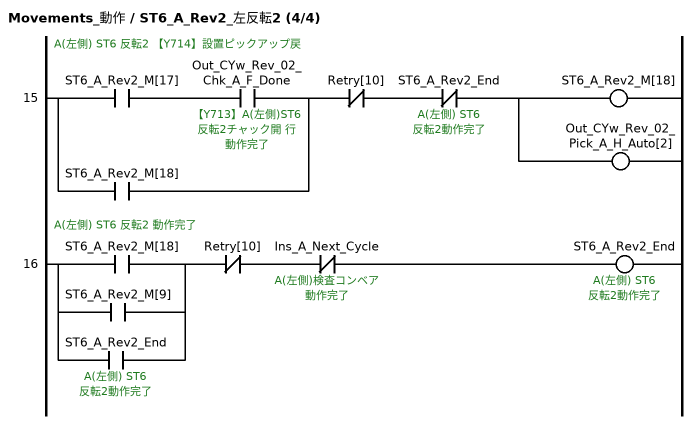
(* [picture p48: Movements_動作 / ST6_A_Rev2_左反転2, rungs 15-16] *)
(* Rung 15: A(左側) ST6 反転2 【Y714】設置ピックアップ戻 *)
_p89 := ((ST6_A_Rev2_M[17] AND Out_CYw_Rev_02_Chk_A_F_Done) OR ST6_A_Rev2_M[18]) AND NOT Retry[10] AND NOT ST6_A_Rev2_End;
ST6_A_Rev2_M[18] := _p89;
Out_CYw_Rev_02_Pick_A_H_Auto[2] := _p89;
(* Rung 16: A(左側) ST6 反転2 動作完了 *)
ST6_A_Rev2_End := (ST6_A_Rev2_M[18] OR ST6_A_Rev2_M[9] OR ST6_A_Rev2_End) AND NOT Retry[10] AND NOT Ins_A_Next_Cycle;

(* Section ST7_A_Dis2_左SF排出: ladder, written here as Structured Text *)

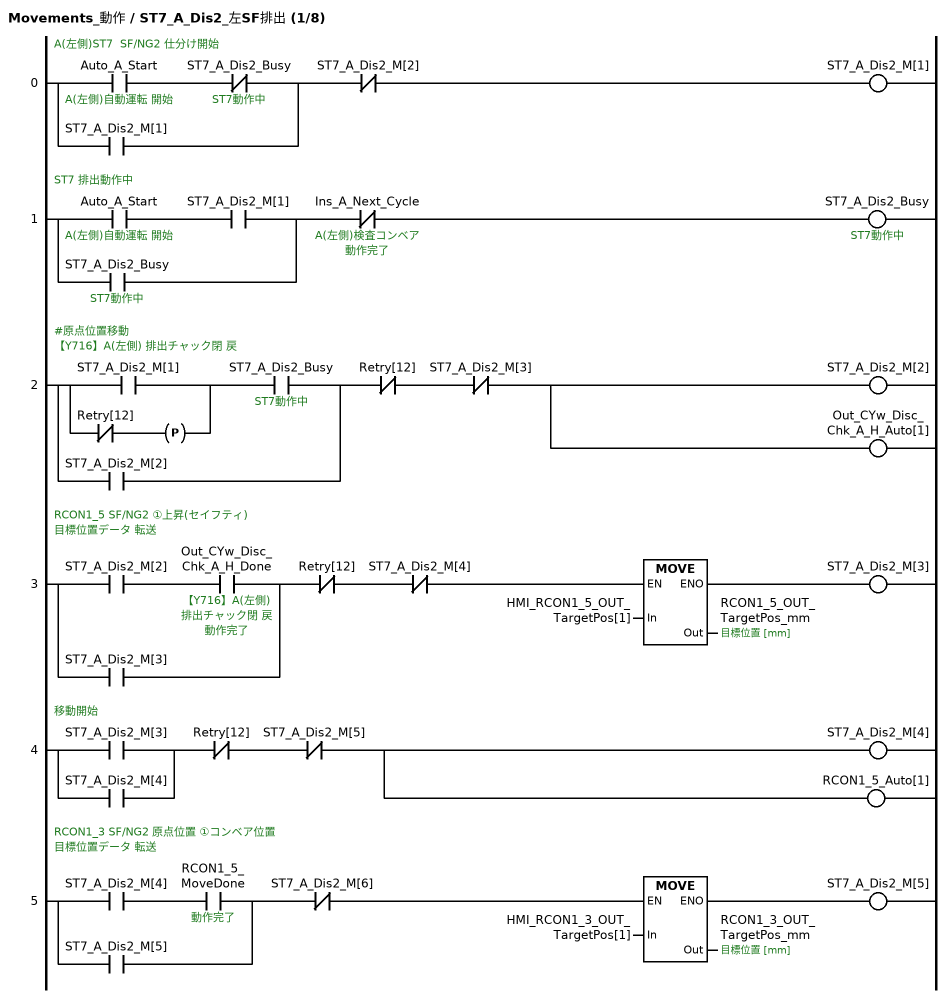
(* Rung 0: A(左側)ST7  SF/NG2 仕分け開始 *)
ST7_A_Dis2_M[1] := ((Auto_A_Start AND NOT ST7_A_Dis2_Busy) OR ST7_A_Dis2_M[1]) AND NOT ST7_A_Dis2_M[2];
(* Rung 1: ST7 排出動作中 *)
ST7_A_Dis2_Busy := ((Auto_A_Start AND ST7_A_Dis2_M[1]) OR ST7_A_Dis2_Busy) AND NOT Ins_A_Next_Cycle;
(* Rung 2: #原点位置移動 / 【Y716】A(左側) 排出チャック閉 戻 *)
_e90(CLK := NOT Retry[12]);
_p91 := (((ST7_A_Dis2_M[1] OR _e90.Q) AND ST7_A_Dis2_Busy) OR ST7_A_Dis2_M[2]) AND NOT Retry[12] AND NOT ST7_A_Dis2_M[3];
ST7_A_Dis2_M[2] := _p91;
Out_CYw_Disc_Chk_A_H_Auto[1] := _p91;
(* Rung 3: RCON1_5 SF/NG2 ①上昇(セイフティ) / 目標位置データ 転送 *)
IF ((ST7_A_Dis2_M[2] AND Out_CYw_Disc_Chk_A_H_Done) OR ST7_A_Dis2_M[3]) AND NOT Retry[12] AND NOT ST7_A_Dis2_M[4] THEN
    RCON1_5_OUT_TargetPos_mm := HMI_RCON1_5_OUT_TargetPos[1];
END_IF;
ST7_A_Dis2_M[3] := ((ST7_A_Dis2_M[2] AND Out_CYw_Disc_Chk_A_H_Done) OR ST7_A_Dis2_M[3]) AND NOT Retry[12] AND NOT ST7_A_Dis2_M[4];
(* Rung 4: 移動開始 *)
_p92 := (ST7_A_Dis2_M[3] OR ST7_A_Dis2_M[4]) AND NOT Retry[12] AND NOT ST7_A_Dis2_M[5];
ST7_A_Dis2_M[4] := _p92;
RCON1_5_Auto[1] := _p92;
(* Rung 5: RCON1_3 SF/NG2 原点位置 ①コンベア位置 / 目標位置データ 転送 *)
IF ((ST7_A_Dis2_M[4] AND RCON1_5_MoveDone) OR ST7_A_Dis2_M[5]) AND NOT ST7_A_Dis2_M[6] THEN
    RCON1_3_OUT_TargetPos_mm := HMI_RCON1_3_OUT_TargetPos[1];
END_IF;
ST7_A_Dis2_M[5] := ((ST7_A_Dis2_M[4] AND RCON1_5_MoveDone) OR ST7_A_Dis2_M[5]) AND NOT ST7_A_Dis2_M[6];

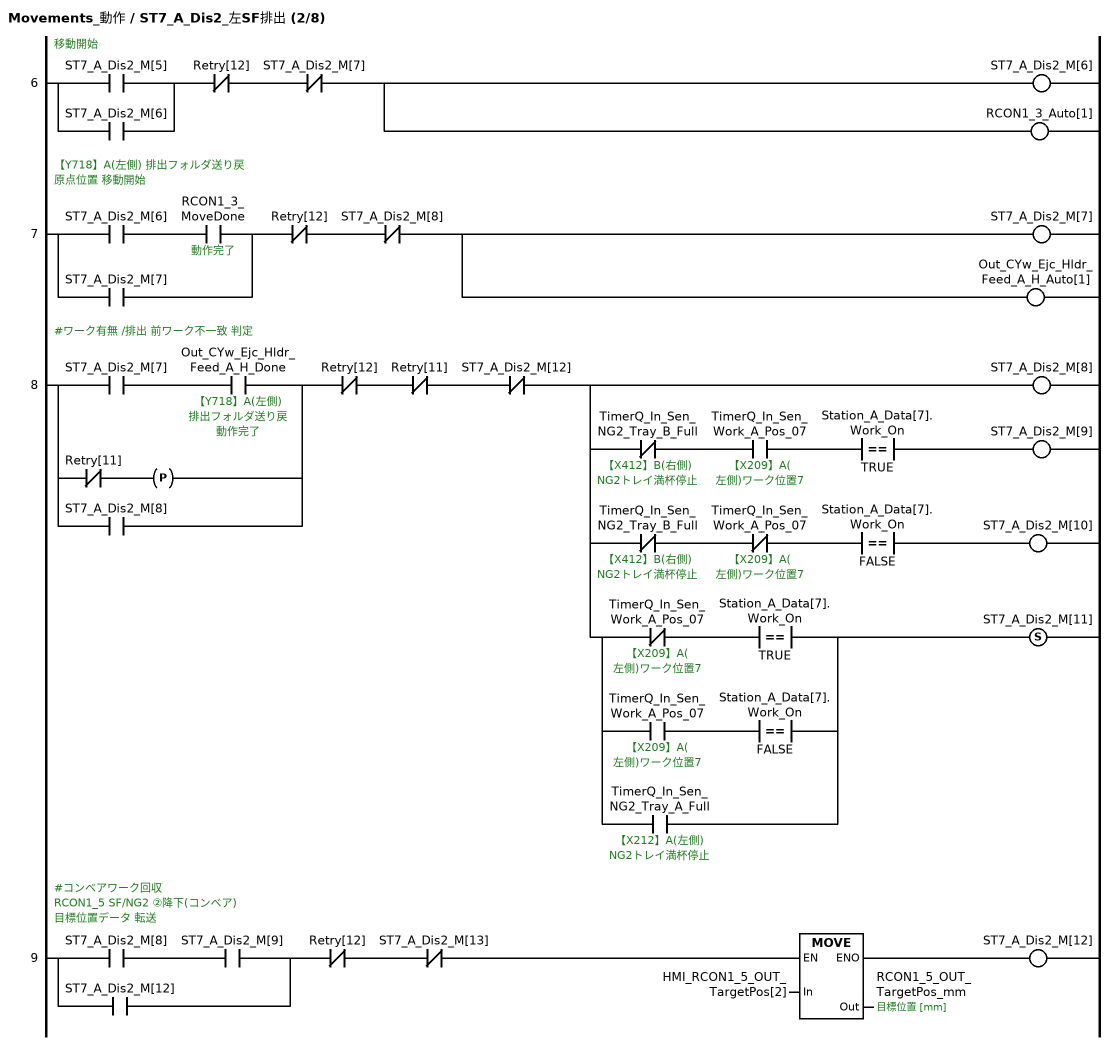
(* Rung 6: 移動開始 *)
_p93 := (ST7_A_Dis2_M[5] OR ST7_A_Dis2_M[6]) AND NOT Retry[12] AND NOT ST7_A_Dis2_M[7];
ST7_A_Dis2_M[6] := _p93;
RCON1_3_Auto[1] := _p93;
(* Rung 7: 【Y718】A(左側) 排出フォルダ送り戻 / 原点位置 移動開始 *)
_p94 := ((ST7_A_Dis2_M[6] AND RCON1_3_MoveDone) OR ST7_A_Dis2_M[7]) AND NOT Retry[12] AND NOT ST7_A_Dis2_M[8];
ST7_A_Dis2_M[7] := _p94;
Out_CYw_Ejc_Hldr_Feed_A_H_Auto[1] := _p94;
(* Rung 8: #ワーク有無 /排出 前ワーク不一致 判定 *)
_e95(CLK := NOT Retry[11]);
_p96 := ((ST7_A_Dis2_M[7] AND Out_CYw_Ejc_Hldr_Feed_A_H_Done) OR _e95.Q OR ST7_A_Dis2_M[8]) AND NOT Retry[12] AND NOT Retry[11] AND NOT ST7_A_Dis2_M[12];
ST7_A_Dis2_M[8] := _p96;
ST7_A_Dis2_M[9] := _p96 AND NOT TimerQ_In_Sen_NG2_Tray_B_Full AND TimerQ_In_Sen_Work_A_Pos_07 AND (Station_A_Data[7].Work_On = TRUE);
ST7_A_Dis2_M[10] := _p96 AND NOT TimerQ_In_Sen_NG2_Tray_B_Full AND NOT TimerQ_In_Sen_Work_A_Pos_07 AND (Station_A_Data[7].Work_On = FALSE);
IF _p96 AND ((NOT TimerQ_In_Sen_Work_A_Pos_07 AND (Station_A_Data[7].Work_On = TRUE)) OR (TimerQ_In_Sen_Work_A_Pos_07 AND (Station_A_Data[7].Work_On = FALSE)) OR TimerQ_In_Sen_NG2_Tray_A_Full) THEN
    ST7_A_Dis2_M[11] := TRUE;
END_IF;
(* Rung 9: #コンベアワーク回収 / RCON1_5 SF/NG2 ②降下(コンベア) / 目標位置データ 転送 *)
IF ((ST7_A_Dis2_M[8] AND ST7_A_Dis2_M[9]) OR ST7_A_Dis2_M[12]) AND NOT Retry[12] AND NOT ST7_A_Dis2_M[13] THEN
    RCON1_5_OUT_TargetPos_mm := HMI_RCON1_5_OUT_TargetPos[2];
END_IF;
ST7_A_Dis2_M[12] := ((ST7_A_Dis2_M[8] AND ST7_A_Dis2_M[9]) OR ST7_A_Dis2_M[12]) AND NOT Retry[12] AND NOT ST7_A_Dis2_M[13];

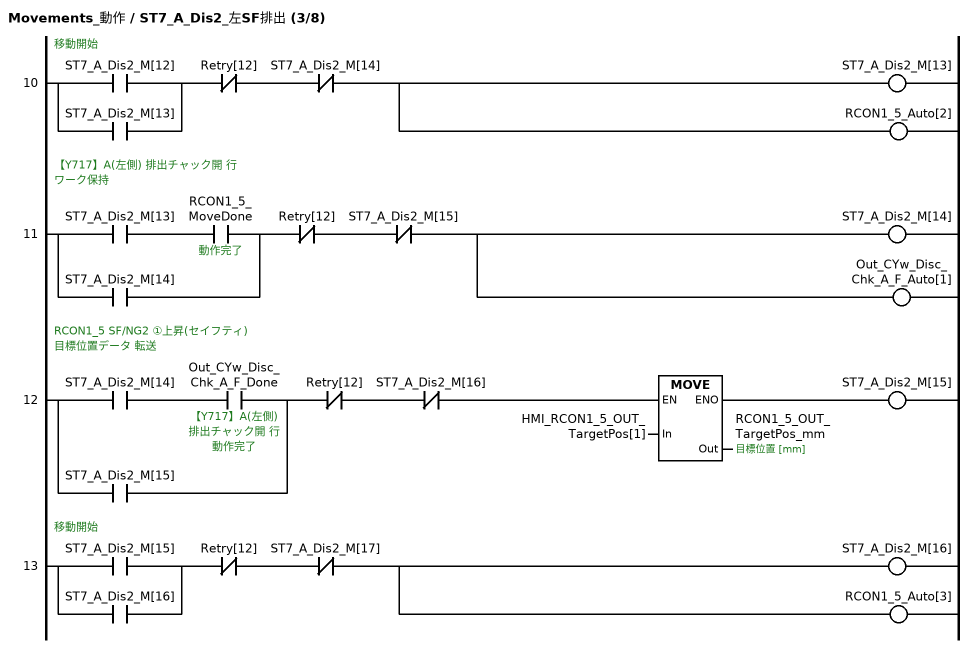
(* Rung 10: 移動開始 *)
_p97 := (ST7_A_Dis2_M[12] OR ST7_A_Dis2_M[13]) AND NOT Retry[12] AND NOT ST7_A_Dis2_M[14];
ST7_A_Dis2_M[13] := _p97;
RCON1_5_Auto[2] := _p97;
(* Rung 11: 【Y717】A(左側) 排出チャック開 行 / ワーク保持 *)
_p98 := ((ST7_A_Dis2_M[13] AND RCON1_5_MoveDone) OR ST7_A_Dis2_M[14]) AND NOT Retry[12] AND NOT ST7_A_Dis2_M[15];
ST7_A_Dis2_M[14] := _p98;
Out_CYw_Disc_Chk_A_F_Auto[1] := _p98;
(* Rung 12: RCON1_5 SF/NG2 ①上昇(セイフティ) / 目標位置データ 転送 *)
IF ((ST7_A_Dis2_M[14] AND Out_CYw_Disc_Chk_A_F_Done) OR ST7_A_Dis2_M[15]) AND NOT Retry[12] AND NOT ST7_A_Dis2_M[16] THEN
    RCON1_5_OUT_TargetPos_mm := HMI_RCON1_5_OUT_TargetPos[1];
END_IF;
ST7_A_Dis2_M[15] := ((ST7_A_Dis2_M[14] AND Out_CYw_Disc_Chk_A_F_Done) OR ST7_A_Dis2_M[15]) AND NOT Retry[12] AND NOT ST7_A_Dis2_M[16];
(* Rung 13: 移動開始 *)
_p99 := (ST7_A_Dis2_M[15] OR ST7_A_Dis2_M[16]) AND NOT Retry[12] AND NOT ST7_A_Dis2_M[17];
ST7_A_Dis2_M[16] := _p99;
RCON1_5_Auto[3] := _p99;

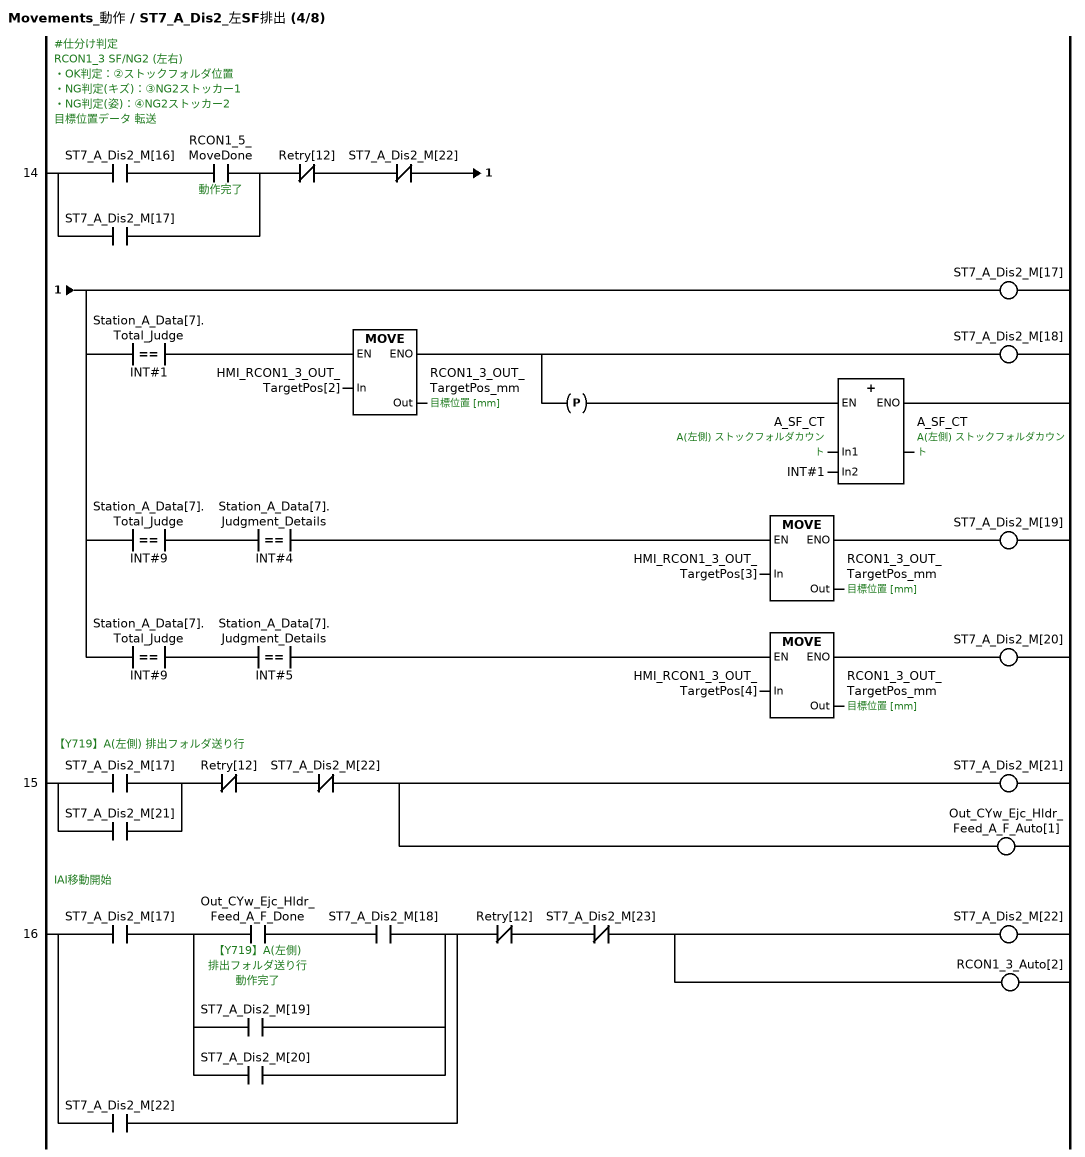
(* Rung 14: #仕分け判定 / RCON1_3 SF/NG2 (左右) / ・OK判定：②ストックフォルダ位置 / ・NG判定(キズ)：③NG2ストッカー1 / ・NG判定(姿)：④NG2ストッカー2 / 目標位置データ 転送 *)
_p100 := ((ST7_A_Dis2_M[16] AND RCON1_5_MoveDone) OR ST7_A_Dis2_M[17]) AND NOT Retry[12] AND NOT ST7_A_Dis2_M[22];
ST7_A_Dis2_M[17] := _p100;
IF _p100 AND (Station_A_Data[7].Total_Judge = INT#1) THEN
    RCON1_3_OUT_TargetPos_mm := HMI_RCON1_3_OUT_TargetPos[2];
END_IF;
_p101 := _p100 AND (Station_A_Data[7].Total_Judge = INT#1);
ST7_A_Dis2_M[18] := _p101;
_e102(CLK := _p101);
IF _e102.Q THEN A_SF_CT := A_SF_CT + INT#1; END_IF;
IF _p100 AND (Station_A_Data[7].Total_Judge = INT#9) AND (Station_A_Data[7].Judgment_Details = INT#4) THEN
    RCON1_3_OUT_TargetPos_mm := HMI_RCON1_3_OUT_TargetPos[3];
END_IF;
ST7_A_Dis2_M[19] := _p100 AND (Station_A_Data[7].Total_Judge = INT#9) AND (Station_A_Data[7].Judgment_Details = INT#4);
IF _p100 AND (Station_A_Data[7].Total_Judge = INT#9) AND (Station_A_Data[7].Judgment_Details = INT#5) THEN
    RCON1_3_OUT_TargetPos_mm := HMI_RCON1_3_OUT_TargetPos[4];
END_IF;
ST7_A_Dis2_M[20] := _p100 AND (Station_A_Data[7].Total_Judge = INT#9) AND (Station_A_Data[7].Judgment_Details = INT#5);
(* Rung 15: 【Y719】A(左側) 排出フォルダ送り行 *)
_p103 := (ST7_A_Dis2_M[17] OR ST7_A_Dis2_M[21]) AND NOT Retry[12] AND NOT ST7_A_Dis2_M[22];
ST7_A_Dis2_M[21] := _p103;
Out_CYw_Ejc_Hldr_Feed_A_F_Auto[1] := _p103;
(* Rung 16: IAI移動開始 *)
_p104 := ((ST7_A_Dis2_M[17] AND ((Out_CYw_Ejc_Hldr_Feed_A_F_Done AND ST7_A_Dis2_M[18]) OR ST7_A_Dis2_M[19] OR ST7_A_Dis2_M[20])) OR ST7_A_Dis2_M[22]) AND NOT Retry[12] AND NOT ST7_A_Dis2_M[23];
ST7_A_Dis2_M[22] := _p104;
RCON1_3_Auto[2] := _p104;

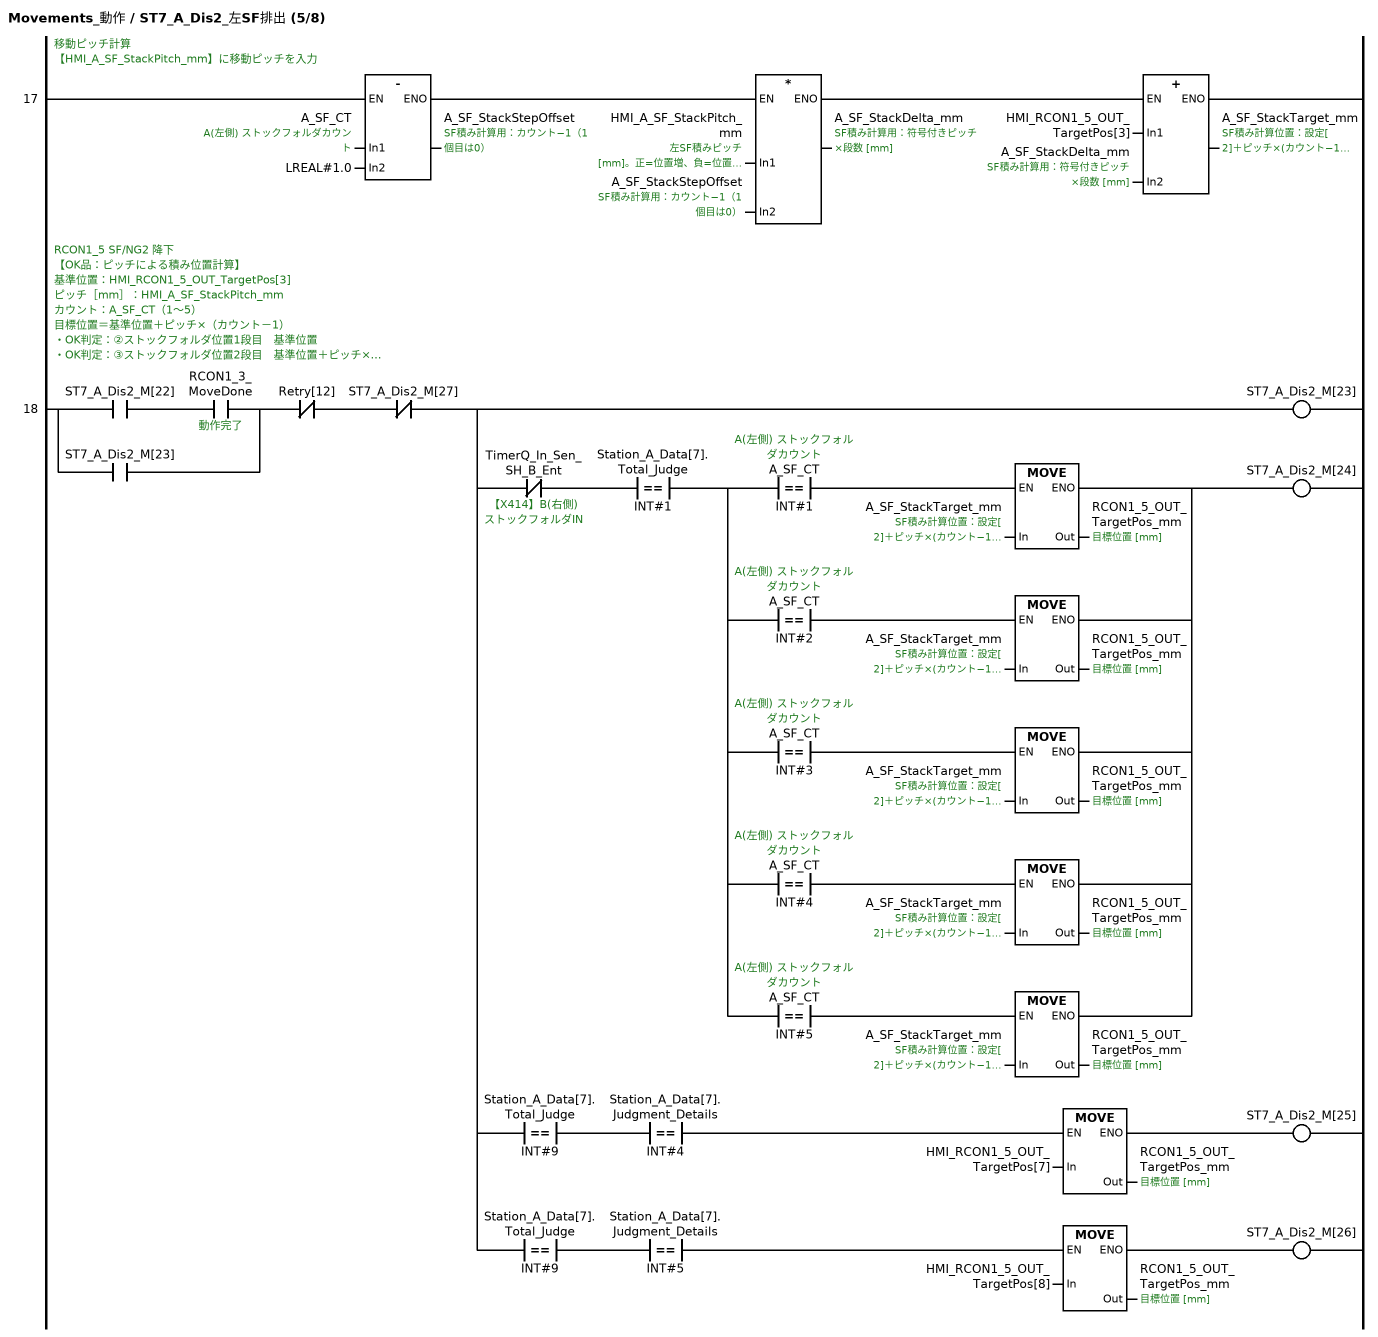
(* Rung 17: 移動ピッチ計算 / 【HMI_A_SF_StackPitch_mm】に移動ピッチを入力 *)
A_SF_StackStepOffset := A_SF_CT - LREAL#1.0;
A_SF_StackDelta_mm := HMI_A_SF_StackPitch_mm * A_SF_StackStepOffset;
A_SF_StackTarget_mm := HMI_RCON1_5_OUT_TargetPos[3] + A_SF_StackDelta_mm;
(* Rung 18: RCON1_5 SF/NG2 降下 / 【OK品：ピッチによる積み位置計算】 / 基準位置：HMI_RCON1_5_OUT_TargetPos[3] / ピッチ［mm］：HMI_A_SF_StackPitch_mm / カウント：A_SF_CT（1～5） / 目標位置＝基準位置＋ピッチ×（カウント－1） / ・OK判定：②ストックフォルダ位置1段目　基準位置 / ・OK判定：③ストックフォルダ位置2段目　基準位置＋ピッチ×1 / ・OK判定：④ストックフォルダ位置3段目　基準位置＋ピッチ×2 / ・OK判定：⑤ストックフォルダ位置4段目　基準位置＋ピッチ×3 / ・OK判定：⑥ストックフォルダ位置5段目　基準位置＋ピッチ×4 / 【NG品：従来の固定位置を使用】 / ・NG判定(キズ)：⑦NG2ストッカー1 / ・NG判定(姿)：⑧NG2ストッカー2 / 目標位置データ 転送 *)
_p105 := ((ST7_A_Dis2_M[22] AND RCON1_3_MoveDone) OR ST7_A_Dis2_M[23]) AND NOT Retry[12] AND NOT ST7_A_Dis2_M[27];
ST7_A_Dis2_M[23] := _p105;
_p106 := _p105 AND NOT TimerQ_In_Sen_SH_B_Ent AND (Station_A_Data[7].Total_Judge = INT#1);
IF _p106 AND (A_SF_CT = INT#1) THEN RCON1_5_OUT_TargetPos_mm := A_SF_StackTarget_mm; END_IF;
IF _p106 AND (A_SF_CT = INT#2) THEN RCON1_5_OUT_TargetPos_mm := A_SF_StackTarget_mm; END_IF;
IF _p106 AND (A_SF_CT = INT#3) THEN RCON1_5_OUT_TargetPos_mm := A_SF_StackTarget_mm; END_IF;
IF _p106 AND (A_SF_CT = INT#4) THEN RCON1_5_OUT_TargetPos_mm := A_SF_StackTarget_mm; END_IF;
IF _p106 AND (A_SF_CT = INT#5) THEN RCON1_5_OUT_TargetPos_mm := A_SF_StackTarget_mm; END_IF;
ST7_A_Dis2_M[24] := _p106 AND ((A_SF_CT = INT#1) OR (A_SF_CT = INT#2) OR (A_SF_CT = INT#3) OR (A_SF_CT = INT#4) OR (A_SF_CT = INT#5));
IF _p105 AND (Station_A_Data[7].Total_Judge = INT#9) AND (Station_A_Data[7].Judgment_Details = INT#4) THEN
    RCON1_5_OUT_TargetPos_mm := HMI_RCON1_5_OUT_TargetPos[7];
END_IF;
ST7_A_Dis2_M[25] := _p105 AND (Station_A_Data[7].Total_Judge = INT#9) AND (Station_A_Data[7].Judgment_Details = INT#4);
IF _p105 AND (Station_A_Data[7].Total_Judge = INT#9) AND (Station_A_Data[7].Judgment_Details = INT#5) THEN
    RCON1_5_OUT_TargetPos_mm := HMI_RCON1_5_OUT_TargetPos[8];
END_IF;
ST7_A_Dis2_M[26] := _p105 AND (Station_A_Data[7].Total_Judge = INT#9) AND (Station_A_Data[7].Judgment_Details = INT#5);

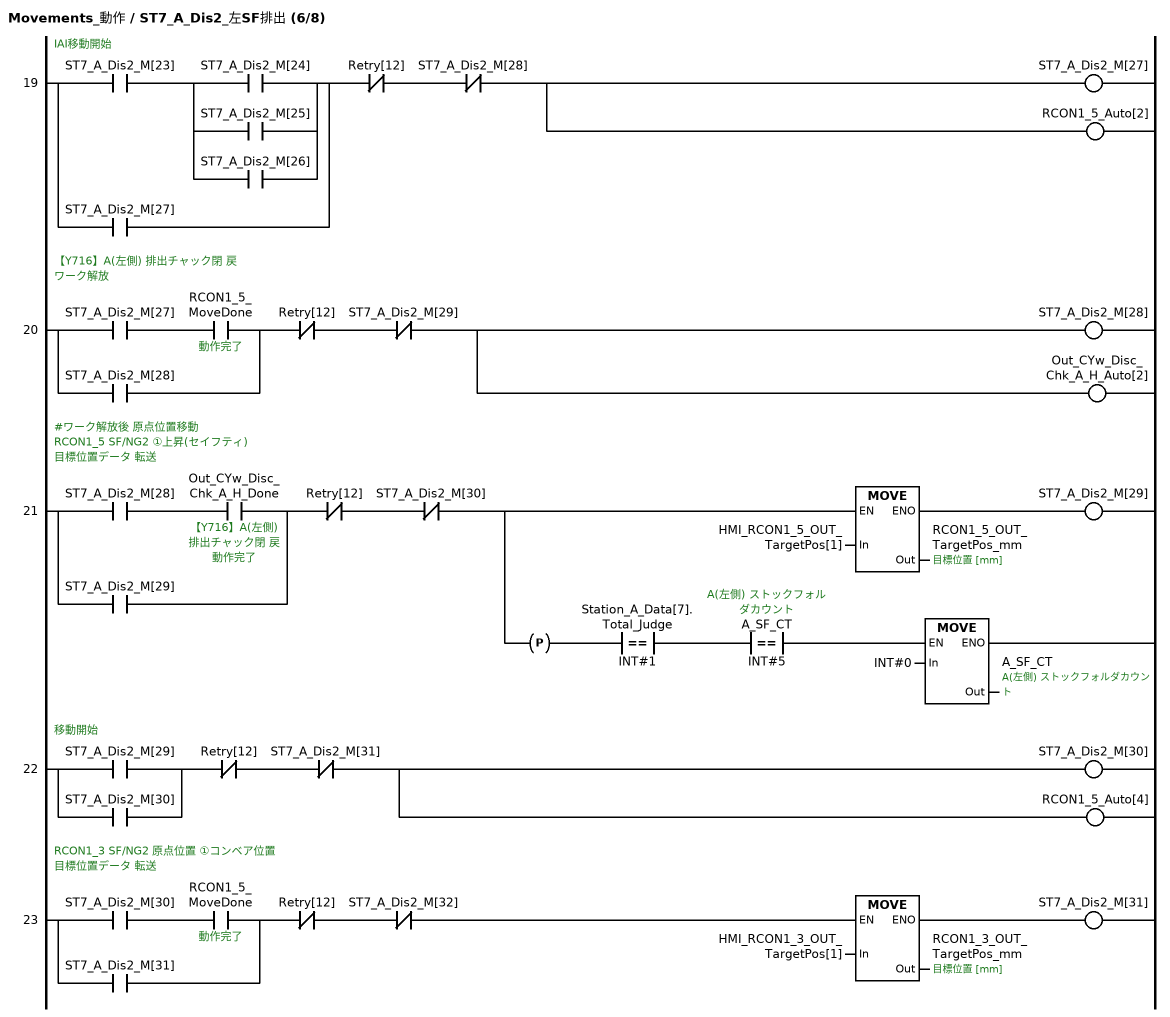
(* Rung 19: IAI移動開始 *)
_p107 := ((ST7_A_Dis2_M[23] AND (ST7_A_Dis2_M[24] OR ST7_A_Dis2_M[25] OR ST7_A_Dis2_M[26])) OR ST7_A_Dis2_M[27]) AND NOT Retry[12] AND NOT ST7_A_Dis2_M[28];
ST7_A_Dis2_M[27] := _p107;
RCON1_5_Auto[2] := _p107;
(* Rung 20: 【Y716】A(左側) 排出チャック閉 戻 / ワーク解放 *)
_p108 := ((ST7_A_Dis2_M[27] AND RCON1_5_MoveDone) OR ST7_A_Dis2_M[28]) AND NOT Retry[12] AND NOT ST7_A_Dis2_M[29];
ST7_A_Dis2_M[28] := _p108;
Out_CYw_Disc_Chk_A_H_Auto[2] := _p108;
(* Rung 21: #ワーク解放後 原点位置移動 / RCON1_5 SF/NG2 ①上昇(セイフティ) / 目標位置データ 転送 *)
_p109 := ((ST7_A_Dis2_M[28] AND Out_CYw_Disc_Chk_A_H_Done) OR ST7_A_Dis2_M[29]) AND NOT Retry[12] AND NOT ST7_A_Dis2_M[30];
IF _p109 THEN RCON1_5_OUT_TargetPos_mm := HMI_RCON1_5_OUT_TargetPos[1]; END_IF;
ST7_A_Dis2_M[29] := _p109;
_e110(CLK := _p109);
IF _e110.Q AND (Station_A_Data[7].Total_Judge = INT#1) AND (A_SF_CT = INT#5) THEN
    A_SF_CT := INT#0;
END_IF;
(* Rung 22: 移動開始 *)
_p111 := (ST7_A_Dis2_M[29] OR ST7_A_Dis2_M[30]) AND NOT Retry[12] AND NOT ST7_A_Dis2_M[31];
ST7_A_Dis2_M[30] := _p111;
RCON1_5_Auto[4] := _p111;
(* Rung 23: RCON1_3 SF/NG2 原点位置 ①コンベア位置 / 目標位置データ 転送 *)
IF ((ST7_A_Dis2_M[30] AND RCON1_5_MoveDone) OR ST7_A_Dis2_M[31]) AND NOT Retry[12] AND NOT ST7_A_Dis2_M[32] THEN
    RCON1_3_OUT_TargetPos_mm := HMI_RCON1_3_OUT_TargetPos[1];
END_IF;
ST7_A_Dis2_M[31] := ((ST7_A_Dis2_M[30] AND RCON1_5_MoveDone) OR ST7_A_Dis2_M[31]) AND NOT Retry[12] AND NOT ST7_A_Dis2_M[32];

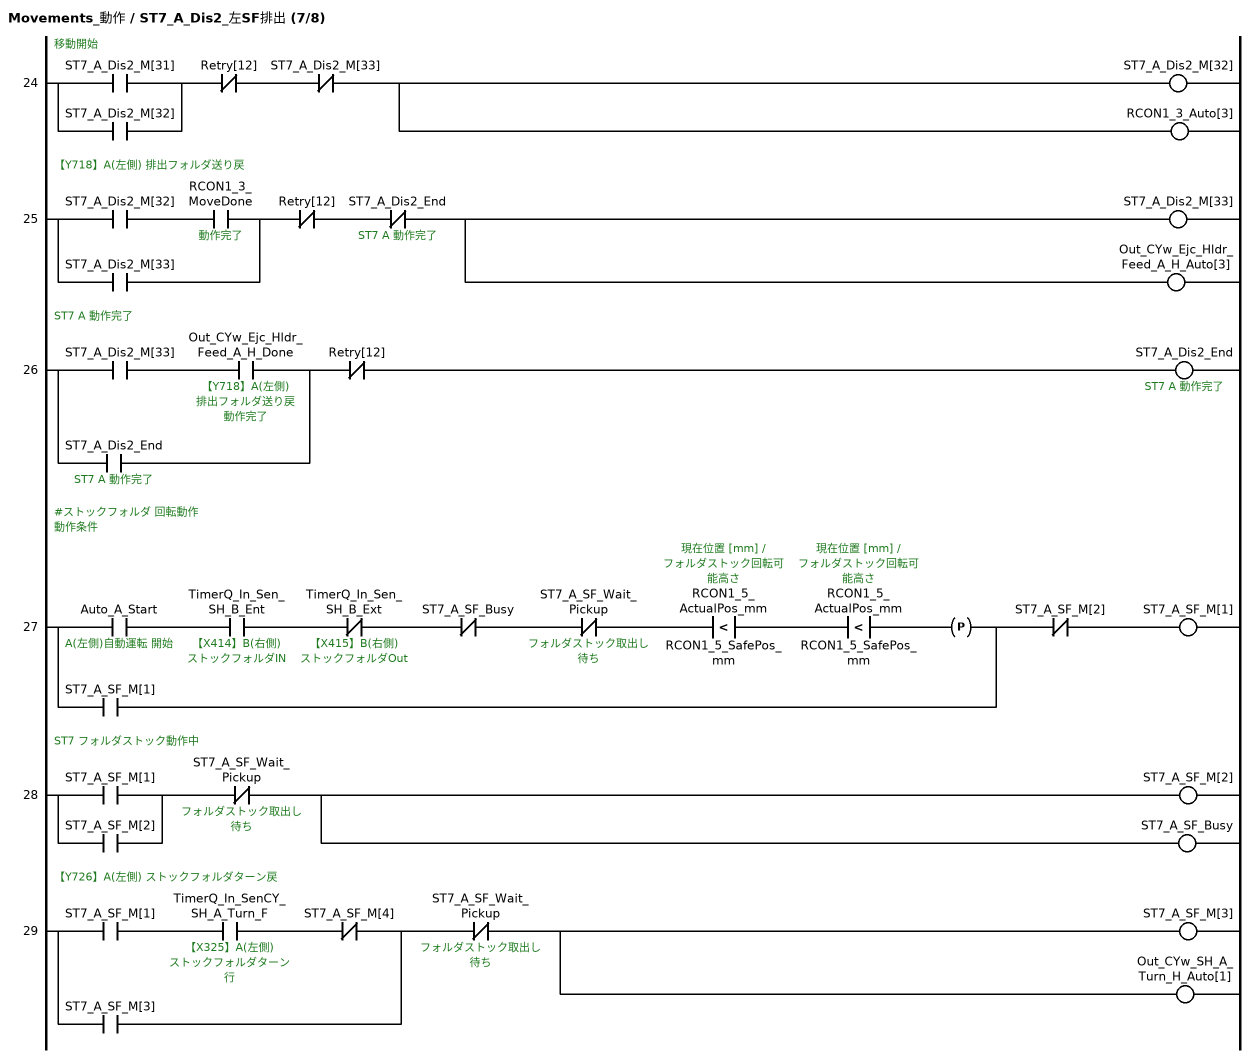
(* Rung 24: 移動開始 *)
_p112 := (ST7_A_Dis2_M[31] OR ST7_A_Dis2_M[32]) AND NOT Retry[12] AND NOT ST7_A_Dis2_M[33];
ST7_A_Dis2_M[32] := _p112;
RCON1_3_Auto[3] := _p112;
(* Rung 25: 【Y718】A(左側) 排出フォルダ送り戻 *)
_p113 := ((ST7_A_Dis2_M[32] AND RCON1_3_MoveDone) OR ST7_A_Dis2_M[33]) AND NOT Retry[12] AND NOT ST7_A_Dis2_End;
ST7_A_Dis2_M[33] := _p113;
Out_CYw_Ejc_Hldr_Feed_A_H_Auto[3] := _p113;
(* Rung 26: ST7 A 動作完了 *)
ST7_A_Dis2_End := ((ST7_A_Dis2_M[33] AND Out_CYw_Ejc_Hldr_Feed_A_H_Done) OR ST7_A_Dis2_End) AND NOT Retry[12];
(* Rung 27: #ストックフォルダ 回転動作 / 動作条件 *)
_e114(CLK := Auto_A_Start AND TimerQ_In_Sen_SH_B_Ent AND NOT TimerQ_In_Sen_SH_B_Ext AND NOT ST7_A_SF_Busy AND NOT ST7_A_SF_Wait_Pickup AND (RCON1_5_ActualPos_mm < RCON1_5_SafePos_mm) AND (RCON1_5_ActualPos_mm < RCON1_5_SafePos_mm));
ST7_A_SF_M[1] := (_e114.Q OR ST7_A_SF_M[1]) AND NOT ST7_A_SF_M[2];
(* Rung 28: ST7 フォルダストック動作中 *)
_p115 := (ST7_A_SF_M[1] OR ST7_A_SF_M[2]) AND NOT ST7_A_SF_Wait_Pickup;
ST7_A_SF_M[2] := _p115;
ST7_A_SF_Busy := _p115;
(* Rung 29: 【Y726】A(左側) ストックフォルダターン戻 *)
_p116 := ((ST7_A_SF_M[1] AND TimerQ_In_SenCY_SH_A_Turn_F AND NOT ST7_A_SF_M[4]) OR ST7_A_SF_M[3]) AND NOT ST7_A_SF_Wait_Pickup;
ST7_A_SF_M[3] := _p116;
Out_CYw_SH_A_Turn_H_Auto[1] := _p116;

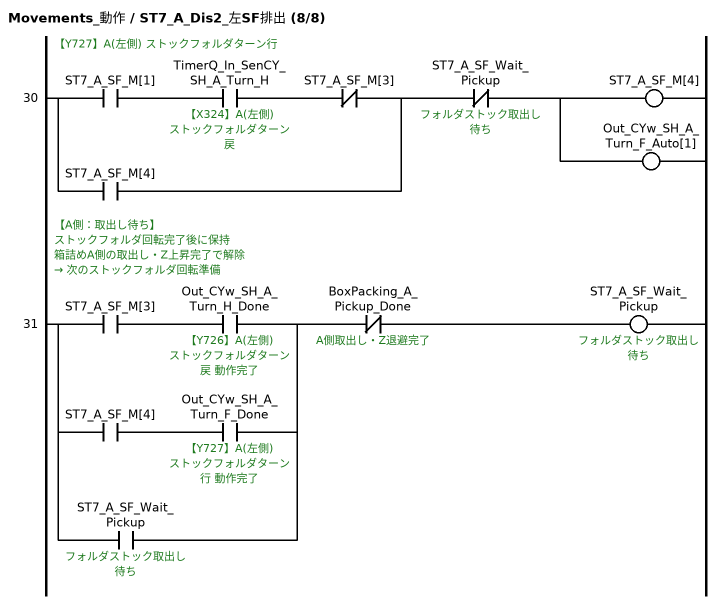
(* Rung 30: 【Y727】A(左側) ストックフォルダターン行 *)
_p117 := ((ST7_A_SF_M[1] AND TimerQ_In_SenCY_SH_A_Turn_H AND NOT ST7_A_SF_M[3]) OR ST7_A_SF_M[4]) AND NOT ST7_A_SF_Wait_Pickup;
ST7_A_SF_M[4] := _p117;
Out_CYw_SH_A_Turn_F_Auto[1] := _p117;
(* Rung 31: 【A側：取出し待ち】 / ストックフォルダ回転完了後に保持 / 箱詰めA側の取出し・Z上昇完了で解除 / → 次のストックフォルダ回転準備 *)
ST7_A_SF_Wait_Pickup := ((ST7_A_SF_M[3] AND Out_CYw_SH_A_Turn_H_Done) OR (ST7_A_SF_M[4] AND Out_CYw_SH_A_Turn_F_Done) OR ST7_A_SF_Wait_Pickup) AND NOT BoxPacking_A_Pickup_Done;

(* Section Destacker_段バラシ: ladder, written here as Structured Text *)

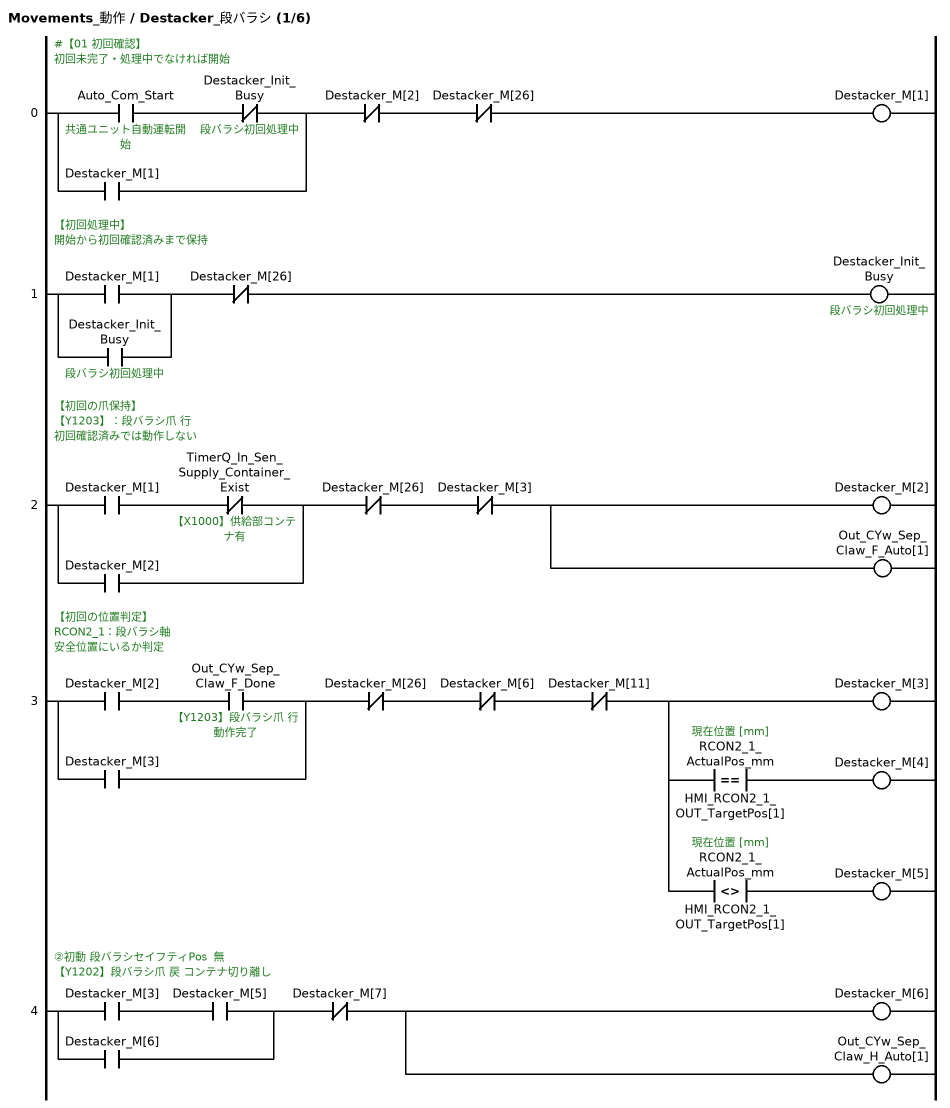
(* Rung 0: #【01 初回確認】 / 初回未完了・処理中でなければ開始 *)
Destacker_M[1] := ((Auto_Com_Start AND NOT Destacker_Init_Busy) OR Destacker_M[1]) AND NOT Destacker_M[2] AND NOT Destacker_M[26];
(* Rung 1: 【初回処理中】 / 開始から初回確認済みまで保持 *)
Destacker_Init_Busy := (Destacker_M[1] OR Destacker_Init_Busy) AND NOT Destacker_M[26];
(* Rung 2: 【初回の爪保持】 / 【Y1203】：段バラシ爪 行 / 初回確認済みでは動作しない *)
_p118 := ((Destacker_M[1] AND NOT TimerQ_In_Sen_Supply_Container_Exist) OR Destacker_M[2]) AND NOT Destacker_M[26] AND NOT Destacker_M[3];
Destacker_M[2] := _p118;
Out_CYw_Sep_Claw_F_Auto[1] := _p118;
(* Rung 3: 【初回の位置判定】 / RCON2_1：段バラシ軸 / 安全位置にいるか判定 *)
_p119 := ((Destacker_M[2] AND Out_CYw_Sep_Claw_F_Done) OR Destacker_M[3]) AND NOT Destacker_M[26] AND NOT Destacker_M[6] AND NOT Destacker_M[11];
Destacker_M[3] := _p119;
Destacker_M[4] := _p119 AND (RCON2_1_ActualPos_mm = HMI_RCON2_1_OUT_TargetPos[1]);
Destacker_M[5] := _p119 AND (RCON2_1_ActualPos_mm <> HMI_RCON2_1_OUT_TargetPos[1]);
(* Rung 4: ②初動 段バラシセイフティPos  無 / 【Y1202】段バラシ爪 戻 コンテナ切り離し *)
_p120 := ((Destacker_M[3] AND Destacker_M[5]) OR Destacker_M[6]) AND NOT Destacker_M[7];
Destacker_M[6] := _p120;
Out_CYw_Sep_Claw_H_Auto[1] := _p120;

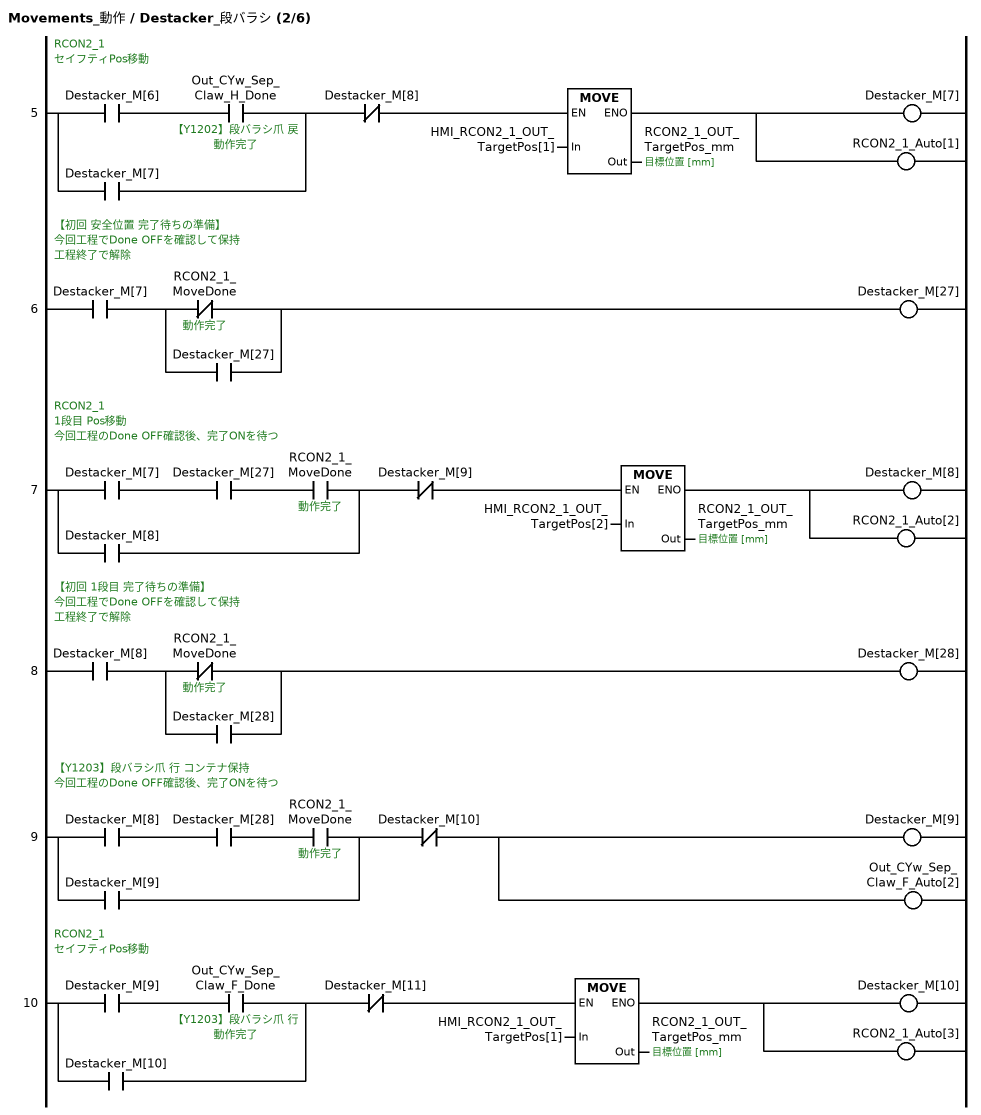
(* Rung 5: RCON2_1 / セイフティPos移動 *)
IF ((Destacker_M[6] AND Out_CYw_Sep_Claw_H_Done) OR Destacker_M[7]) AND NOT Destacker_M[8] THEN
    RCON2_1_OUT_TargetPos_mm := HMI_RCON2_1_OUT_TargetPos[1];
END_IF;
_p121 := ((Destacker_M[6] AND Out_CYw_Sep_Claw_H_Done) OR Destacker_M[7]) AND NOT Destacker_M[8];
Destacker_M[7] := _p121;
RCON2_1_Auto[1] := _p121;
(* Rung 6: 【初回 安全位置 完了待ちの準備】 / 今回工程でDone OFFを確認して保持 / 工程終了で解除 *)
Destacker_M[27] := Destacker_M[7] AND (NOT RCON2_1_MoveDone OR Destacker_M[27]);
(* Rung 7: RCON2_1 / 1段目 Pos移動 / 今回工程のDone OFF確認後、完了ONを待つ *)
IF ((Destacker_M[7] AND Destacker_M[27] AND RCON2_1_MoveDone) OR Destacker_M[8]) AND NOT Destacker_M[9] THEN
    RCON2_1_OUT_TargetPos_mm := HMI_RCON2_1_OUT_TargetPos[2];
END_IF;
_p122 := ((Destacker_M[7] AND Destacker_M[27] AND RCON2_1_MoveDone) OR Destacker_M[8]) AND NOT Destacker_M[9];
Destacker_M[8] := _p122;
RCON2_1_Auto[2] := _p122;
(* Rung 8: 【初回 1段目 完了待ちの準備】 / 今回工程でDone OFFを確認して保持 / 工程終了で解除 *)
Destacker_M[28] := Destacker_M[8] AND (NOT RCON2_1_MoveDone OR Destacker_M[28]);
(* Rung 9: 【Y1203】段バラシ爪 行 コンテナ保持 / 今回工程のDone OFF確認後、完了ONを待つ *)
_p123 := ((Destacker_M[8] AND Destacker_M[28] AND RCON2_1_MoveDone) OR Destacker_M[9]) AND NOT Destacker_M[10];
Destacker_M[9] := _p123;
Out_CYw_Sep_Claw_F_Auto[2] := _p123;
(* Rung 10: RCON2_1 / セイフティPos移動 *)
IF ((Destacker_M[9] AND Out_CYw_Sep_Claw_F_Done) OR Destacker_M[10]) AND NOT Destacker_M[11] THEN
    RCON2_1_OUT_TargetPos_mm := HMI_RCON2_1_OUT_TargetPos[1];
END_IF;
_p124 := ((Destacker_M[9] AND Out_CYw_Sep_Claw_F_Done) OR Destacker_M[10]) AND NOT Destacker_M[11];
Destacker_M[10] := _p124;
RCON2_1_Auto[3] := _p124;

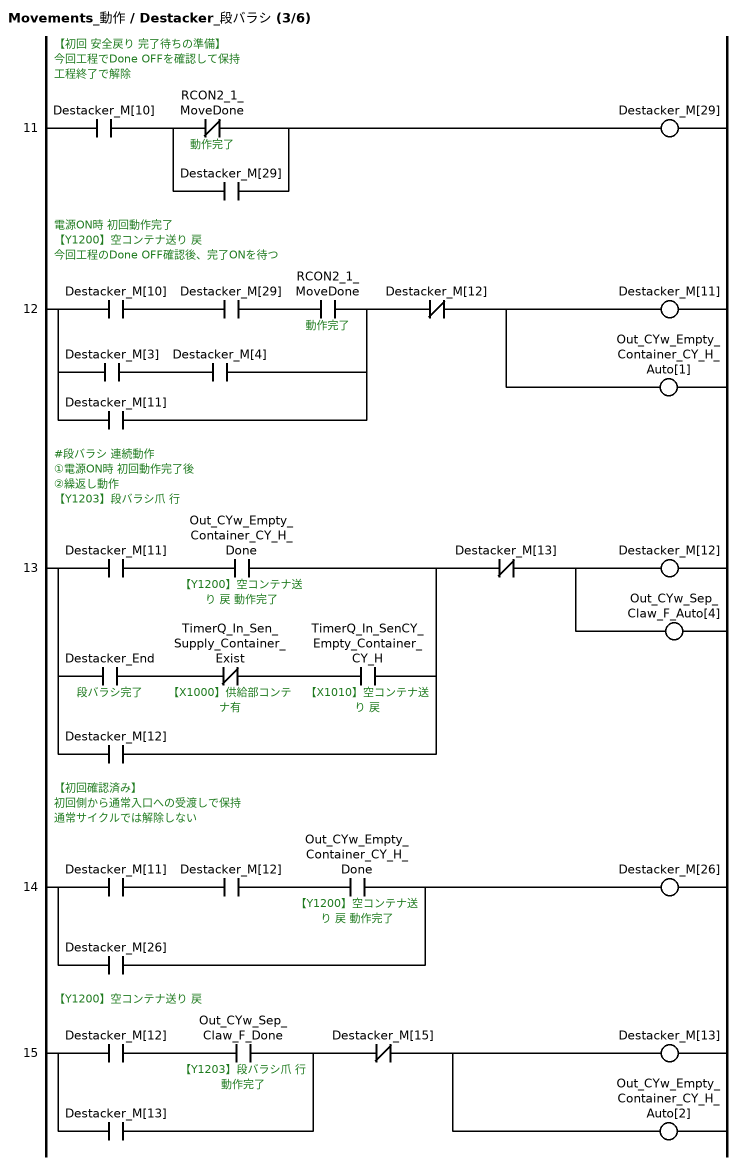
(* Rung 11: 【初回 安全戻り 完了待ちの準備】 / 今回工程でDone OFFを確認して保持 / 工程終了で解除 *)
Destacker_M[29] := Destacker_M[10] AND (NOT RCON2_1_MoveDone OR Destacker_M[29]);
(* Rung 12: 電源ON時 初回動作完了 / 【Y1200】空コンテナ送り 戻 / 今回工程のDone OFF確認後、完了ONを待つ *)
_p125 := ((Destacker_M[10] AND Destacker_M[29] AND RCON2_1_MoveDone) OR (Destacker_M[3] AND Destacker_M[4]) OR Destacker_M[11]) AND NOT Destacker_M[12];
Destacker_M[11] := _p125;
Out_CYw_Empty_Container_CY_H_Auto[1] := _p125;
(* Rung 13: #段バラシ 連続動作 / ①電源ON時 初回動作完了後 / ②繰返し動作 / 【Y1203】段バラシ爪 行 *)
_p126 := ((Destacker_M[11] AND Out_CYw_Empty_Container_CY_H_Done) OR (Destacker_End AND NOT TimerQ_In_Sen_Supply_Container_Exist AND TimerQ_In_SenCY_Empty_Container_CY_H) OR Destacker_M[12]) AND NOT Destacker_M[13];
Destacker_M[12] := _p126;
Out_CYw_Sep_Claw_F_Auto[4] := _p126;
(* Rung 14: 【初回確認済み】 / 初回側から通常入口への受渡しで保持 / 通常サイクルでは解除しない *)
Destacker_M[26] := (Destacker_M[11] AND Destacker_M[12] AND Out_CYw_Empty_Container_CY_H_Done) OR Destacker_M[26];
(* Rung 15: 【Y1200】空コンテナ送り 戻 *)
_p127 := ((Destacker_M[12] AND Out_CYw_Sep_Claw_F_Done) OR Destacker_M[13]) AND NOT Destacker_M[15];
Destacker_M[13] := _p127;
Out_CYw_Empty_Container_CY_H_Auto[2] := _p127;

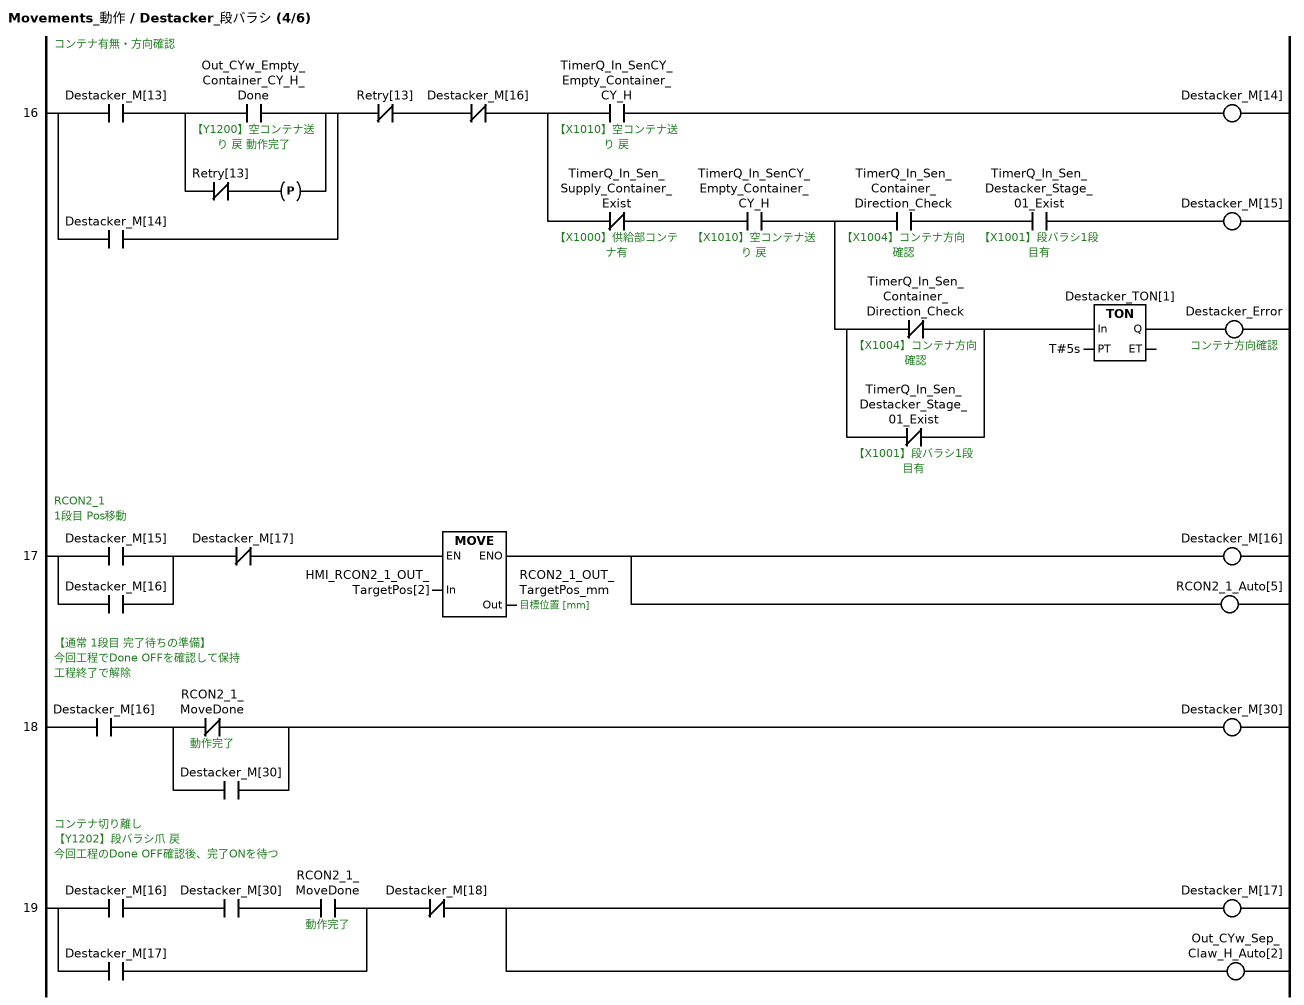
(* Rung 16: コンテナ有無・方向確認 *)
_e128(CLK := Destacker_M[13] AND NOT Retry[13]);
_p129 := ((Destacker_M[13] AND Out_CYw_Empty_Container_CY_H_Done) OR _e128.Q OR Destacker_M[14]) AND NOT Retry[13] AND NOT Destacker_M[16];
Destacker_M[14] := _p129 AND TimerQ_In_SenCY_Empty_Container_CY_H;
_p130 := _p129 AND NOT TimerQ_In_Sen_Supply_Container_Exist AND TimerQ_In_SenCY_Empty_Container_CY_H;
Destacker_M[15] := _p130 AND TimerQ_In_Sen_Container_Direction_Check AND TimerQ_In_Sen_Destacker_Stage_01_Exist;
Destacker_TON[1](In := _p130 AND (NOT TimerQ_In_Sen_Container_Direction_Check OR NOT TimerQ_In_Sen_Destacker_Stage_01_Exist), PT := T#5s);
Destacker_Error := Destacker_TON[1].Q;
(* Rung 17: RCON2_1 / 1段目 Pos移動 *)
IF (Destacker_M[15] OR Destacker_M[16]) AND NOT Destacker_M[17] THEN
    RCON2_1_OUT_TargetPos_mm := HMI_RCON2_1_OUT_TargetPos[2];
END_IF;
_p131 := (Destacker_M[15] OR Destacker_M[16]) AND NOT Destacker_M[17];
Destacker_M[16] := _p131;
RCON2_1_Auto[5] := _p131;
(* Rung 18: 【通常 1段目 完了待ちの準備】 / 今回工程でDone OFFを確認して保持 / 工程終了で解除 *)
Destacker_M[30] := Destacker_M[16] AND (NOT RCON2_1_MoveDone OR Destacker_M[30]);
(* Rung 19: コンテナ切り離し / 【Y1202】段バラシ爪 戻 / 今回工程のDone OFF確認後、完了ONを待つ *)
_p132 := ((Destacker_M[16] AND Destacker_M[30] AND RCON2_1_MoveDone) OR Destacker_M[17]) AND NOT Destacker_M[18];
Destacker_M[17] := _p132;
Out_CYw_Sep_Claw_H_Auto[2] := _p132;

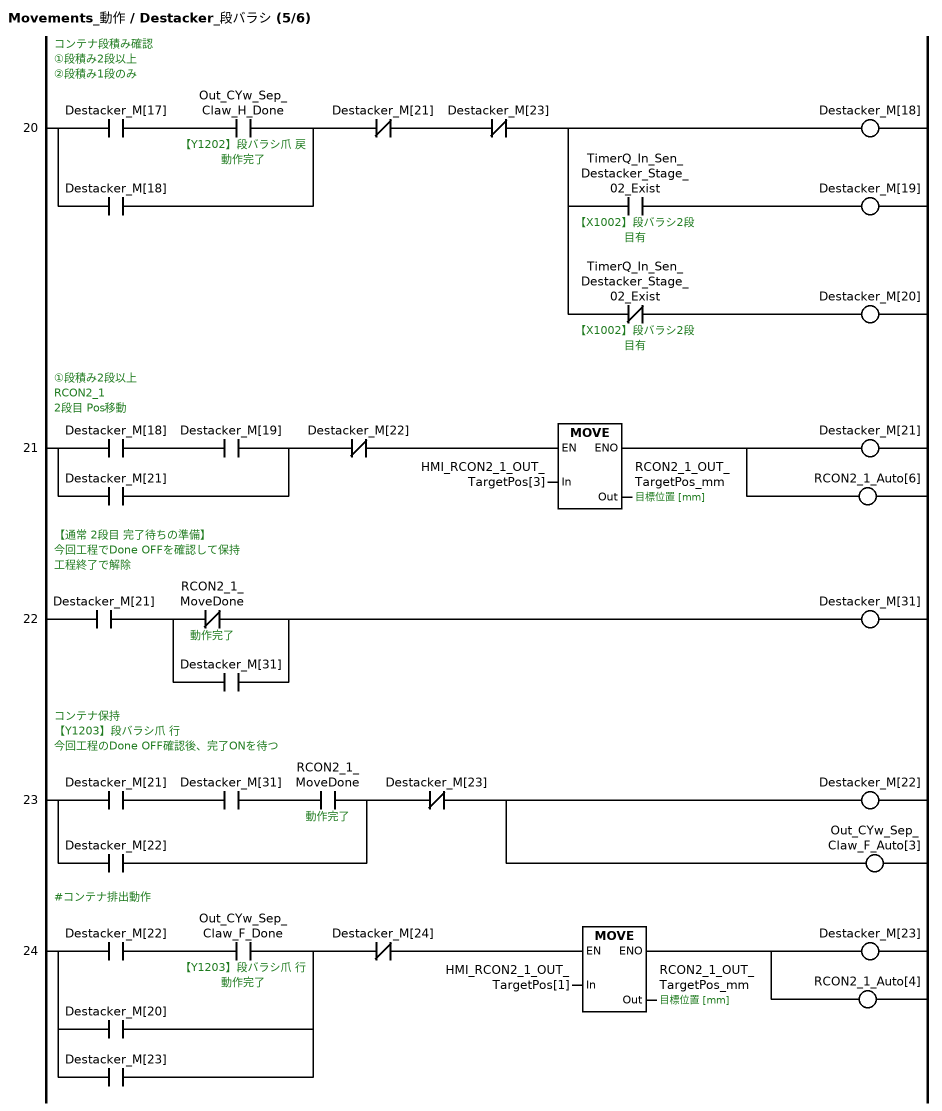
(* Rung 20: コンテナ段積み確認 / ①段積み2段以上 / ②段積み1段のみ *)
_p133 := ((Destacker_M[17] AND Out_CYw_Sep_Claw_H_Done) OR Destacker_M[18]) AND NOT Destacker_M[21] AND NOT Destacker_M[23];
Destacker_M[18] := _p133;
Destacker_M[19] := _p133 AND TimerQ_In_Sen_Destacker_Stage_02_Exist;
Destacker_M[20] := _p133 AND NOT TimerQ_In_Sen_Destacker_Stage_02_Exist;
(* Rung 21: ①段積み2段以上 / RCON2_1 / 2段目 Pos移動 *)
IF ((Destacker_M[18] AND Destacker_M[19]) OR Destacker_M[21]) AND NOT Destacker_M[22] THEN
    RCON2_1_OUT_TargetPos_mm := HMI_RCON2_1_OUT_TargetPos[3];
END_IF;
_p134 := ((Destacker_M[18] AND Destacker_M[19]) OR Destacker_M[21]) AND NOT Destacker_M[22];
Destacker_M[21] := _p134;
RCON2_1_Auto[6] := _p134;
(* Rung 22: 【通常 2段目 完了待ちの準備】 / 今回工程でDone OFFを確認して保持 / 工程終了で解除 *)
Destacker_M[31] := Destacker_M[21] AND (NOT RCON2_1_MoveDone OR Destacker_M[31]);
(* Rung 23: コンテナ保持 / 【Y1203】段バラシ爪 行 / 今回工程のDone OFF確認後、完了ONを待つ *)
_p135 := ((Destacker_M[21] AND Destacker_M[31] AND RCON2_1_MoveDone) OR Destacker_M[22]) AND NOT Destacker_M[23];
Destacker_M[22] := _p135;
Out_CYw_Sep_Claw_F_Auto[3] := _p135;
(* Rung 24: #コンテナ排出動作 *)
IF ((Destacker_M[22] AND Out_CYw_Sep_Claw_F_Done) OR Destacker_M[20] OR Destacker_M[23]) AND NOT Destacker_M[24] THEN
    RCON2_1_OUT_TargetPos_mm := HMI_RCON2_1_OUT_TargetPos[1];
END_IF;
_p136 := ((Destacker_M[22] AND Out_CYw_Sep_Claw_F_Done) OR Destacker_M[20] OR Destacker_M[23]) AND NOT Destacker_M[24];
Destacker_M[23] := _p136;
RCON2_1_Auto[4] := _p136;

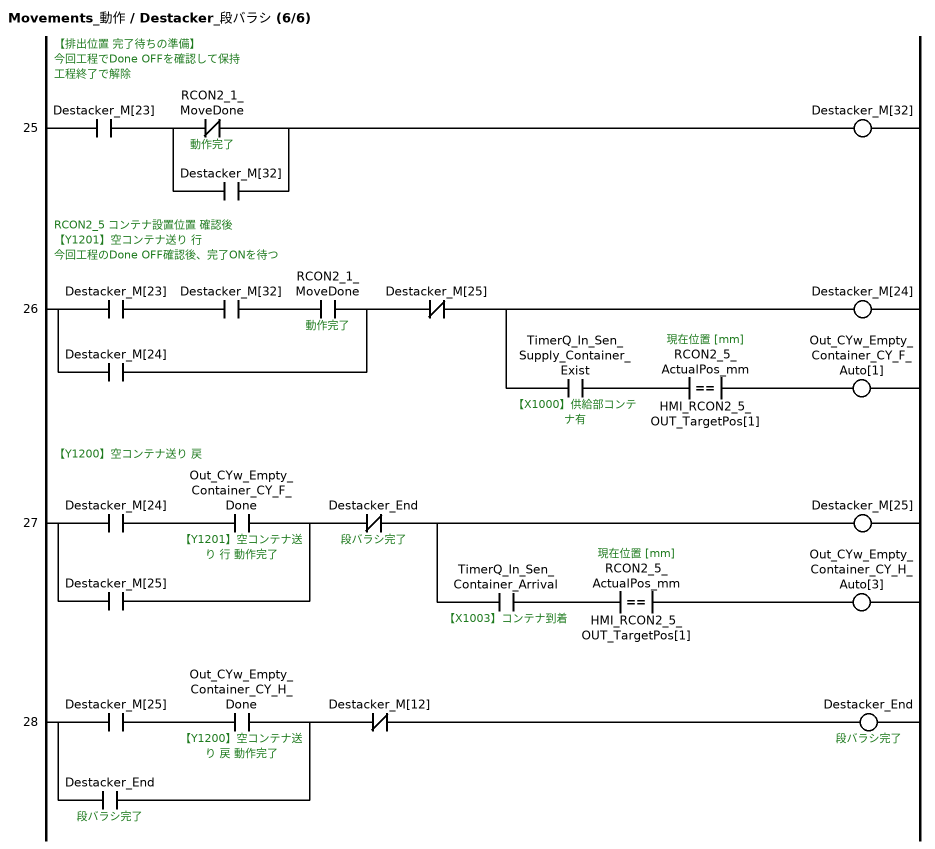
(* Rung 25: 【排出位置 完了待ちの準備】 / 今回工程でDone OFFを確認して保持 / 工程終了で解除 *)
Destacker_M[32] := Destacker_M[23] AND (NOT RCON2_1_MoveDone OR Destacker_M[32]);
(* Rung 26: RCON2_5 コンテナ設置位置 確認後 / 【Y1201】空コンテナ送り 行 / 今回工程のDone OFF確認後、完了ONを待つ *)
_p137 := ((Destacker_M[23] AND Destacker_M[32] AND RCON2_1_MoveDone) OR Destacker_M[24]) AND NOT Destacker_M[25];
Destacker_M[24] := _p137;
Out_CYw_Empty_Container_CY_F_Auto[1] := _p137 AND TimerQ_In_Sen_Supply_Container_Exist AND (RCON2_5_ActualPos_mm = HMI_RCON2_5_OUT_TargetPos[1]);
(* Rung 27: 【Y1200】空コンテナ送り 戻 *)
_p138 := ((Destacker_M[24] AND Out_CYw_Empty_Container_CY_F_Done) OR Destacker_M[25]) AND NOT Destacker_End;
Destacker_M[25] := _p138;
Out_CYw_Empty_Container_CY_H_Auto[3] := _p138 AND TimerQ_In_Sen_Container_Arrival AND (RCON2_5_ActualPos_mm = HMI_RCON2_5_OUT_TargetPos[1]);
(* Rung 28 *)
Destacker_End := ((Destacker_M[25] AND Out_CYw_Empty_Container_CY_H_Done) OR Destacker_End) AND NOT Destacker_M[12];

(* Section BoxPacking_箱詰め: ladder, written here as Structured Text *)

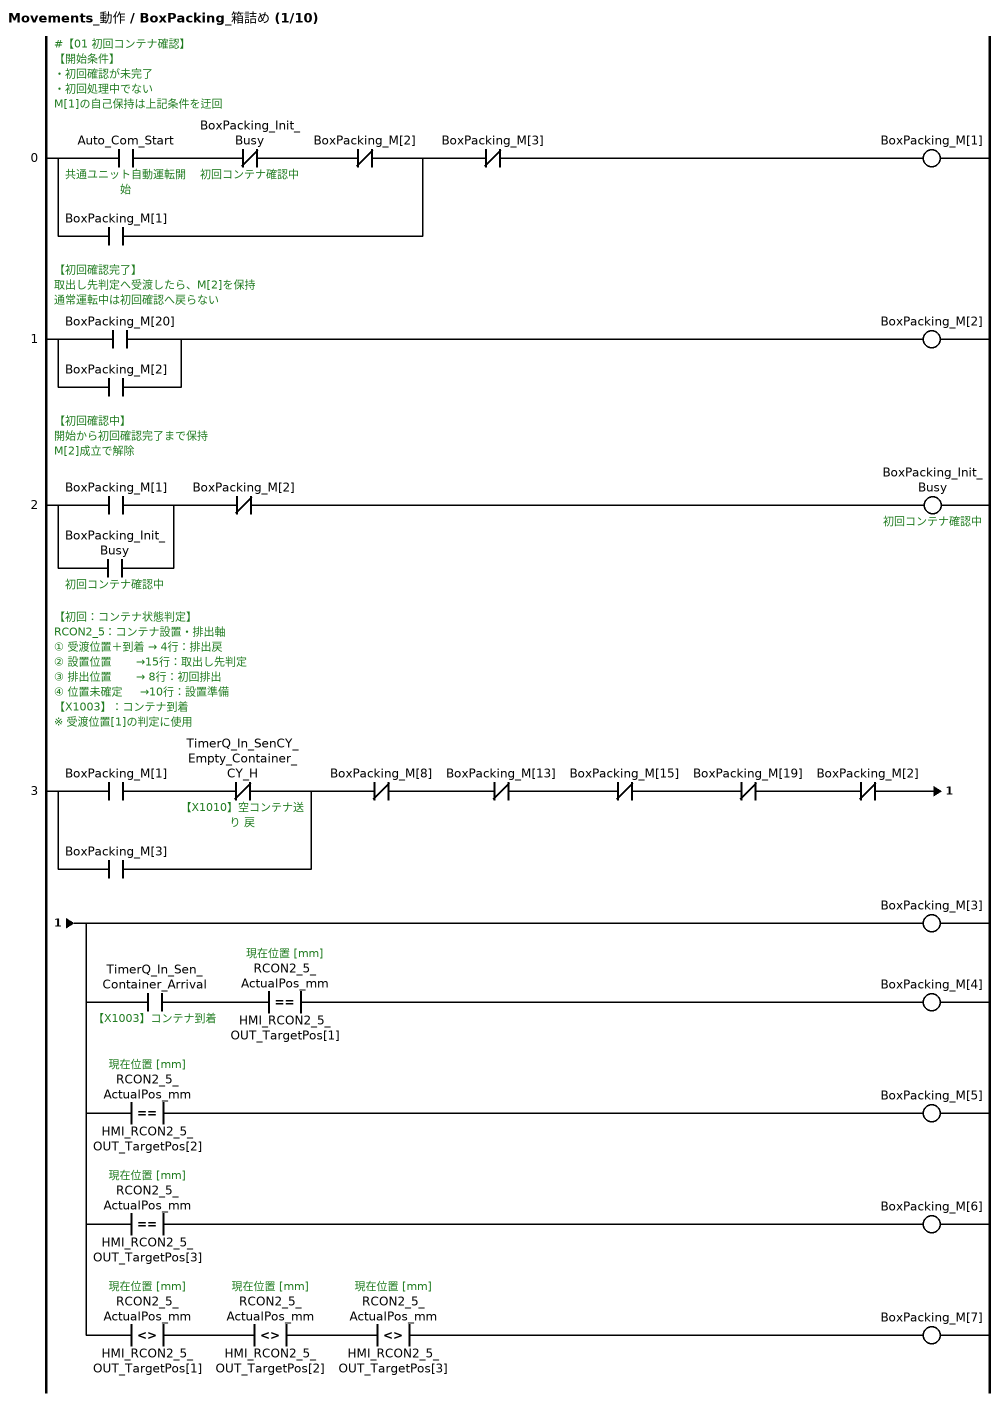
(* Rung 0: #【01 初回コンテナ確認】 / 【開始条件】 / ・初回確認が未完了 / ・初回処理中でない / M[1]の自己保持は上記条件を迂回 *)
BoxPacking_M[1] := ((Auto_Com_Start AND NOT BoxPacking_Init_Busy AND NOT BoxPacking_M[2]) OR BoxPacking_M[1]) AND NOT BoxPacking_M[3];
(* Rung 1: 【初回確認完了】 / 取出し先判定へ受渡したら、M[2]を保持 / 通常運転中は初回確認へ戻らない *)
BoxPacking_M[2] := BoxPacking_M[20] OR BoxPacking_M[2];
(* Rung 2: 【初回確認中】 / 開始から初回確認完了まで保持 / M[2]成立で解除 *)
BoxPacking_Init_Busy := (BoxPacking_M[1] OR BoxPacking_Init_Busy) AND NOT BoxPacking_M[2];
(* Rung 3: 【初回：コンテナ状態判定】 / RCON2_5：コンテナ設置・排出軸 / ① 受渡位置＋到着 → 4行：排出戻 / ② 設置位置       →15行：取出し先判定 / ③ 排出位置       → 8行：初回排出 / ④ 位置未確定     →10行：設置準備 / 【X1003】：コンテナ到着 / ※ 受渡位置[1]の判定に使用 *)
_p139 := ((BoxPacking_M[1] AND NOT TimerQ_In_SenCY_Empty_Container_CY_H) OR BoxPacking_M[3]) AND NOT BoxPacking_M[8] AND NOT BoxPacking_M[13] AND NOT BoxPacking_M[15] AND NOT BoxPacking_M[19] AND NOT BoxPacking_M[2];
BoxPacking_M[3] := _p139;
BoxPacking_M[4] := _p139 AND TimerQ_In_Sen_Container_Arrival AND (RCON2_5_ActualPos_mm = HMI_RCON2_5_OUT_TargetPos[1]);
BoxPacking_M[5] := _p139 AND (RCON2_5_ActualPos_mm = HMI_RCON2_5_OUT_TargetPos[2]);
BoxPacking_M[6] := _p139 AND (RCON2_5_ActualPos_mm = HMI_RCON2_5_OUT_TargetPos[3]);
BoxPacking_M[7] := _p139 AND (RCON2_5_ActualPos_mm <> HMI_RCON2_5_OUT_TargetPos[1]) AND (RCON2_5_ActualPos_mm <> HMI_RCON2_5_OUT_TargetPos[2]) AND (RCON2_5_ActualPos_mm <> HMI_RCON2_5_OUT_TargetPos[3]);

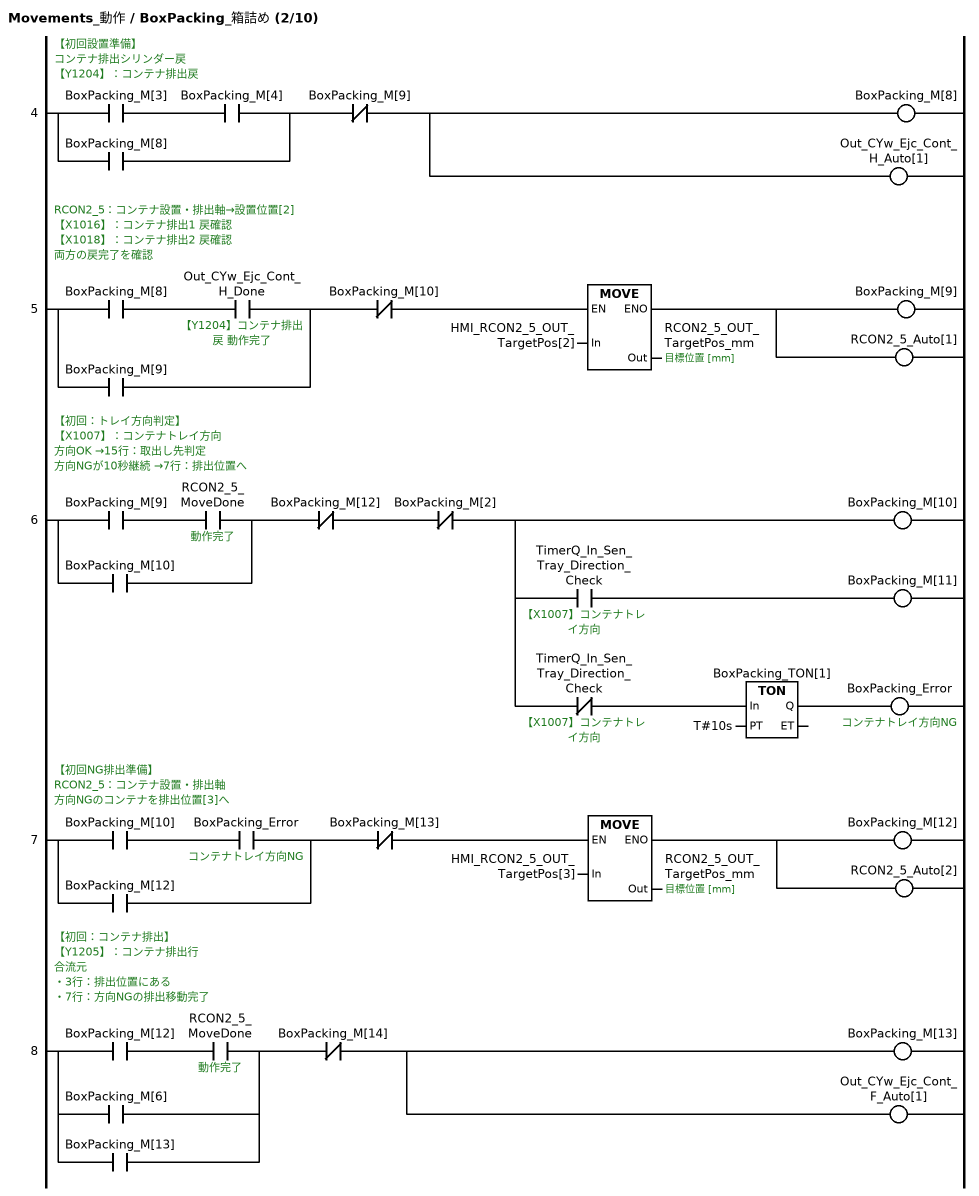
(* Rung 4: 【初回設置準備】 / コンテナ排出シリンダー戻 / 【Y1204】：コンテナ排出戻 *)
_p140 := ((BoxPacking_M[3] AND BoxPacking_M[4]) OR BoxPacking_M[8]) AND NOT BoxPacking_M[9];
BoxPacking_M[8] := _p140;
Out_CYw_Ejc_Cont_H_Auto[1] := _p140;
(* Rung 5: RCON2_5：コンテナ設置・排出軸→設置位置[2] / 【X1016】：コンテナ排出1 戻確認 / 【X1018】：コンテナ排出2 戻確認 / 両方の戻完了を確認 *)
IF ((BoxPacking_M[8] AND Out_CYw_Ejc_Cont_H_Done) OR BoxPacking_M[9]) AND NOT BoxPacking_M[10] THEN
    RCON2_5_OUT_TargetPos_mm := HMI_RCON2_5_OUT_TargetPos[2];
END_IF;
_p141 := ((BoxPacking_M[8] AND Out_CYw_Ejc_Cont_H_Done) OR BoxPacking_M[9]) AND NOT BoxPacking_M[10];
BoxPacking_M[9] := _p141;
RCON2_5_Auto[1] := _p141;
(* Rung 6: 【初回：トレイ方向判定】 / 【X1007】：コンテナトレイ方向 / 方向OK →15行：取出し先判定 / 方向NGが10秒継続 →7行：排出位置へ *)
_p142 := ((BoxPacking_M[9] AND RCON2_5_MoveDone) OR BoxPacking_M[10]) AND NOT BoxPacking_M[12] AND NOT BoxPacking_M[2];
BoxPacking_M[10] := _p142;
BoxPacking_M[11] := _p142 AND TimerQ_In_Sen_Tray_Direction_Check;
BoxPacking_TON[1](In := _p142 AND NOT TimerQ_In_Sen_Tray_Direction_Check, PT := T#10s);
BoxPacking_Error := BoxPacking_TON[1].Q;
(* Rung 7: 【初回NG排出準備】 / RCON2_5：コンテナ設置・排出軸 / 方向NGのコンテナを排出位置[3]へ *)
IF ((BoxPacking_M[10] AND BoxPacking_Error) OR BoxPacking_M[12]) AND NOT BoxPacking_M[13] THEN
    RCON2_5_OUT_TargetPos_mm := HMI_RCON2_5_OUT_TargetPos[3];
END_IF;
_p143 := ((BoxPacking_M[10] AND BoxPacking_Error) OR BoxPacking_M[12]) AND NOT BoxPacking_M[13];
BoxPacking_M[12] := _p143;
RCON2_5_Auto[2] := _p143;
(* Rung 8: 【初回：コンテナ排出】 / 【Y1205】：コンテナ排出行 / 合流元 / ・3行：排出位置にある / ・7行：方向NGの排出移動完了 *)
_p144 := ((BoxPacking_M[12] AND RCON2_5_MoveDone) OR BoxPacking_M[6] OR BoxPacking_M[13]) AND NOT BoxPacking_M[14];
BoxPacking_M[13] := _p144;
Out_CYw_Ejc_Cont_F_Auto[1] := _p144;

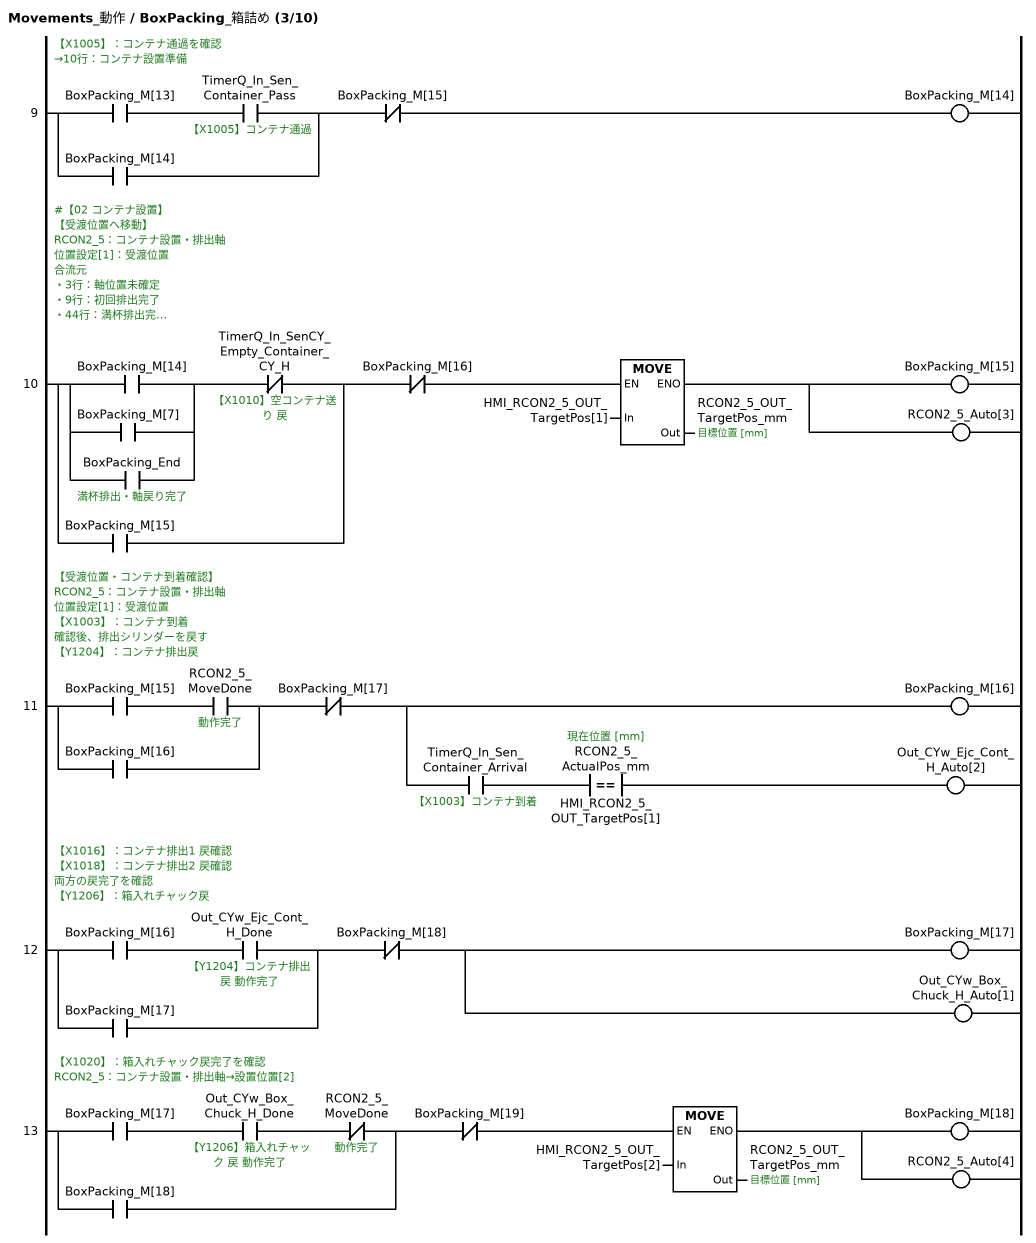
(* Rung 9: 【X1005】：コンテナ通過を確認 / →10行：コンテナ設置準備 *)
BoxPacking_M[14] := ((BoxPacking_M[13] AND TimerQ_In_Sen_Container_Pass) OR BoxPacking_M[14]) AND NOT BoxPacking_M[15];
(* Rung 10: #【02 コンテナ設置】 / 【受渡位置へ移動】 / RCON2_5：コンテナ設置・排出軸 / 位置設定[1]：受渡位置 / 合流元 / ・3行：軸位置未確定 / ・9行：初回排出完了 / ・44行：満杯排出完了 / 44行からは、下記入力のOFFで復帰 / 【X1010】：空コンテナ送り戻確認 *)
IF (((BoxPacking_M[14] OR BoxPacking_M[7] OR BoxPacking_End) AND NOT TimerQ_In_SenCY_Empty_Container_CY_H) OR BoxPacking_M[15]) AND NOT BoxPacking_M[16] THEN
    RCON2_5_OUT_TargetPos_mm := HMI_RCON2_5_OUT_TargetPos[1];
END_IF;
_p145 := (((BoxPacking_M[14] OR BoxPacking_M[7] OR BoxPacking_End) AND NOT TimerQ_In_SenCY_Empty_Container_CY_H) OR BoxPacking_M[15]) AND NOT BoxPacking_M[16];
BoxPacking_M[15] := _p145;
RCON2_5_Auto[3] := _p145;
(* Rung 11: 【受渡位置・コンテナ到着確認】 / RCON2_5：コンテナ設置・排出軸 / 位置設定[1]：受渡位置 / 【X1003】：コンテナ到着 / 確認後、排出シリンダーを戻す / 【Y1204】：コンテナ排出戻 *)
_p146 := ((BoxPacking_M[15] AND RCON2_5_MoveDone) OR BoxPacking_M[16]) AND NOT BoxPacking_M[17];
BoxPacking_M[16] := _p146;
Out_CYw_Ejc_Cont_H_Auto[2] := _p146 AND TimerQ_In_Sen_Container_Arrival AND (RCON2_5_ActualPos_mm = HMI_RCON2_5_OUT_TargetPos[1]);
(* Rung 12: 【X1016】：コンテナ排出1 戻確認 / 【X1018】：コンテナ排出2 戻確認 / 両方の戻完了を確認 / 【Y1206】：箱入れチャック戻 *)
_p147 := ((BoxPacking_M[16] AND Out_CYw_Ejc_Cont_H_Done) OR BoxPacking_M[17]) AND NOT BoxPacking_M[18];
BoxPacking_M[17] := _p147;
Out_CYw_Box_Chuck_H_Auto[1] := _p147;
(* Rung 13: 【X1020】：箱入れチャック戻完了を確認 / RCON2_5：コンテナ設置・排出軸→設置位置[2] *)
IF ((BoxPacking_M[17] AND Out_CYw_Box_Chuck_H_Done AND NOT RCON2_5_MoveDone) OR BoxPacking_M[18]) AND NOT BoxPacking_M[19] THEN
    RCON2_5_OUT_TargetPos_mm := HMI_RCON2_5_OUT_TargetPos[2];
END_IF;
_p148 := ((BoxPacking_M[17] AND Out_CYw_Box_Chuck_H_Done AND NOT RCON2_5_MoveDone) OR BoxPacking_M[18]) AND NOT BoxPacking_M[19];
BoxPacking_M[18] := _p148;
RCON2_5_Auto[4] := _p148;

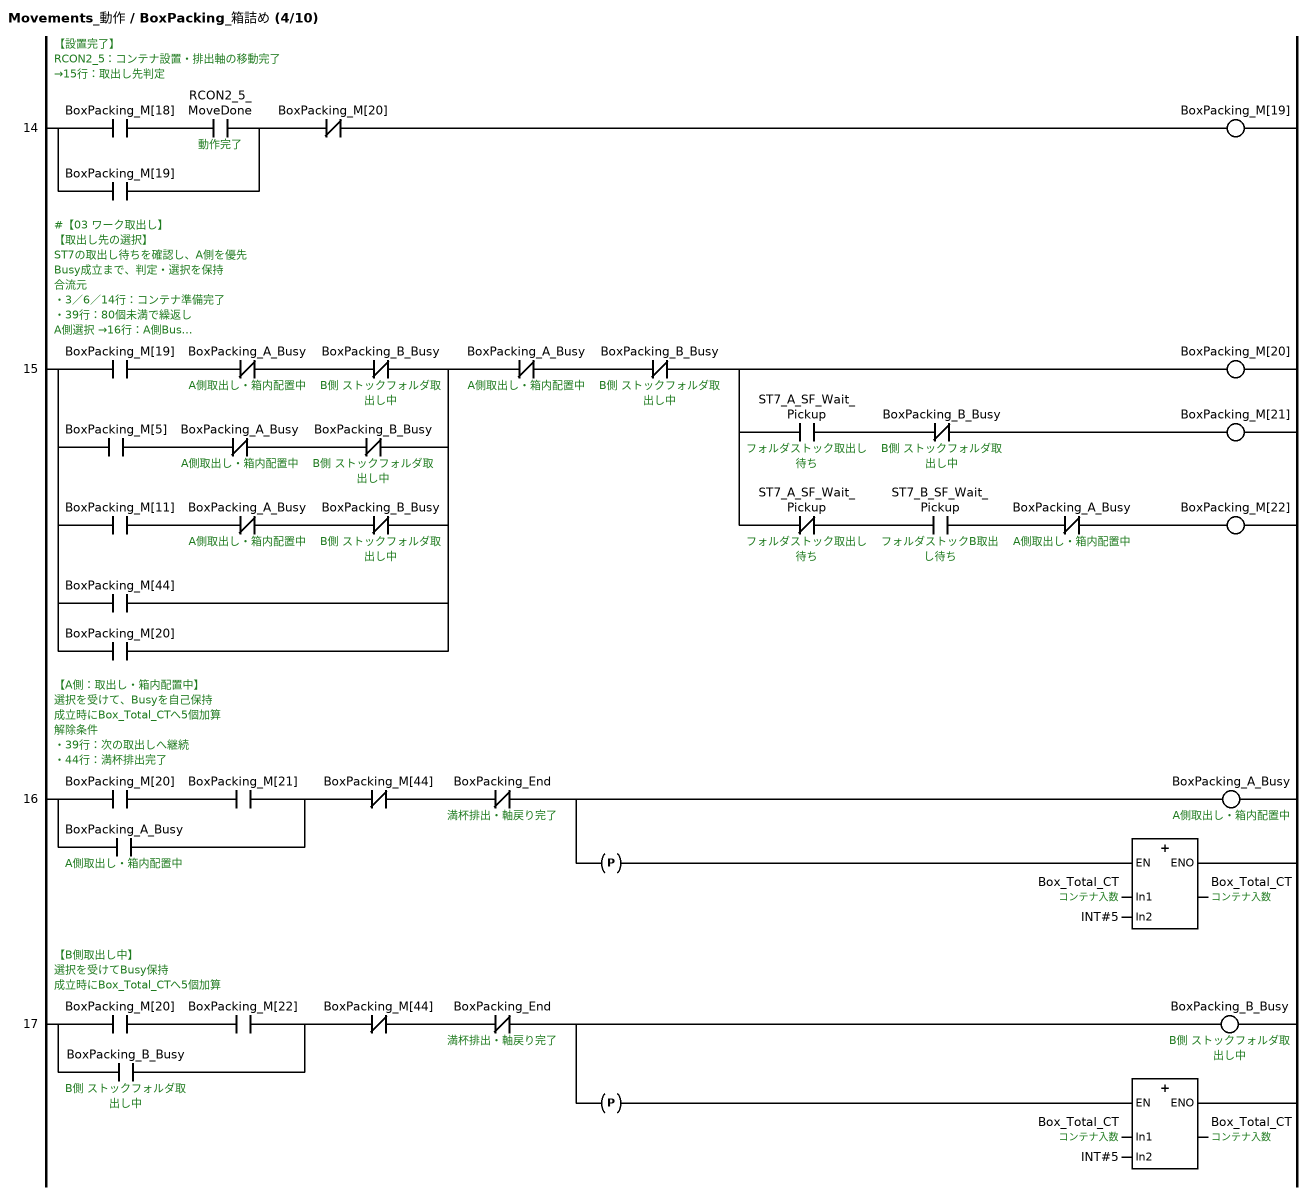
(* Rung 14: 【設置完了】 / RCON2_5：コンテナ設置・排出軸の移動完了 / →15行：取出し先判定 *)
BoxPacking_M[19] := ((BoxPacking_M[18] AND RCON2_5_MoveDone) OR BoxPacking_M[19]) AND NOT BoxPacking_M[20];
(* Rung 15: #【03 ワーク取出し】 / 【取出し先の選択】 / ST7の取出し待ちを確認し、A側を優先 / Busy成立まで、判定・選択を保持 / 合流元 / ・3／6／14行：コンテナ準備完了 / ・39行：80個未満で繰返し / A側選択 →16行：A側Busy / B側選択 →17行：B側Busy *)
_p149 := ((BoxPacking_M[19] AND NOT BoxPacking_A_Busy AND NOT BoxPacking_B_Busy) OR (BoxPacking_M[5] AND NOT BoxPacking_A_Busy AND NOT BoxPacking_B_Busy) OR (BoxPacking_M[11] AND NOT BoxPacking_A_Busy AND NOT BoxPacking_B_Busy) OR BoxPacking_M[44] OR BoxPacking_M[20]) AND NOT BoxPacking_A_Busy AND NOT BoxPacking_B_Busy;
BoxPacking_M[20] := _p149;
BoxPacking_M[21] := _p149 AND ST7_A_SF_Wait_Pickup AND NOT BoxPacking_B_Busy;
BoxPacking_M[22] := _p149 AND NOT ST7_A_SF_Wait_Pickup AND ST7_B_SF_Wait_Pickup AND NOT BoxPacking_A_Busy;
(* Rung 16: 【A側：取出し・箱内配置中】 / 選択を受けて、Busyを自己保持 / 成立時にBox_Total_CTへ5個加算 / 解除条件 / ・39行：次の取出しへ継続 / ・44行：満杯排出完了 *)
_p150 := ((BoxPacking_M[20] AND BoxPacking_M[21]) OR BoxPacking_A_Busy) AND NOT BoxPacking_M[44] AND NOT BoxPacking_End;
BoxPacking_A_Busy := _p150;
_e151(CLK := _p150);
IF _e151.Q THEN Box_Total_CT := Box_Total_CT + INT#5; END_IF;
(* Rung 17: 【B側取出し中】 / 選択を受けてBusy保持 / 成立時にBox_Total_CTへ5個加算 *)
_p152 := ((BoxPacking_M[20] AND BoxPacking_M[22]) OR BoxPacking_B_Busy) AND NOT BoxPacking_M[44] AND NOT BoxPacking_End;
BoxPacking_B_Busy := _p152;
_e153(CLK := _p152);
IF _e153.Q THEN Box_Total_CT := Box_Total_CT + INT#5; END_IF;

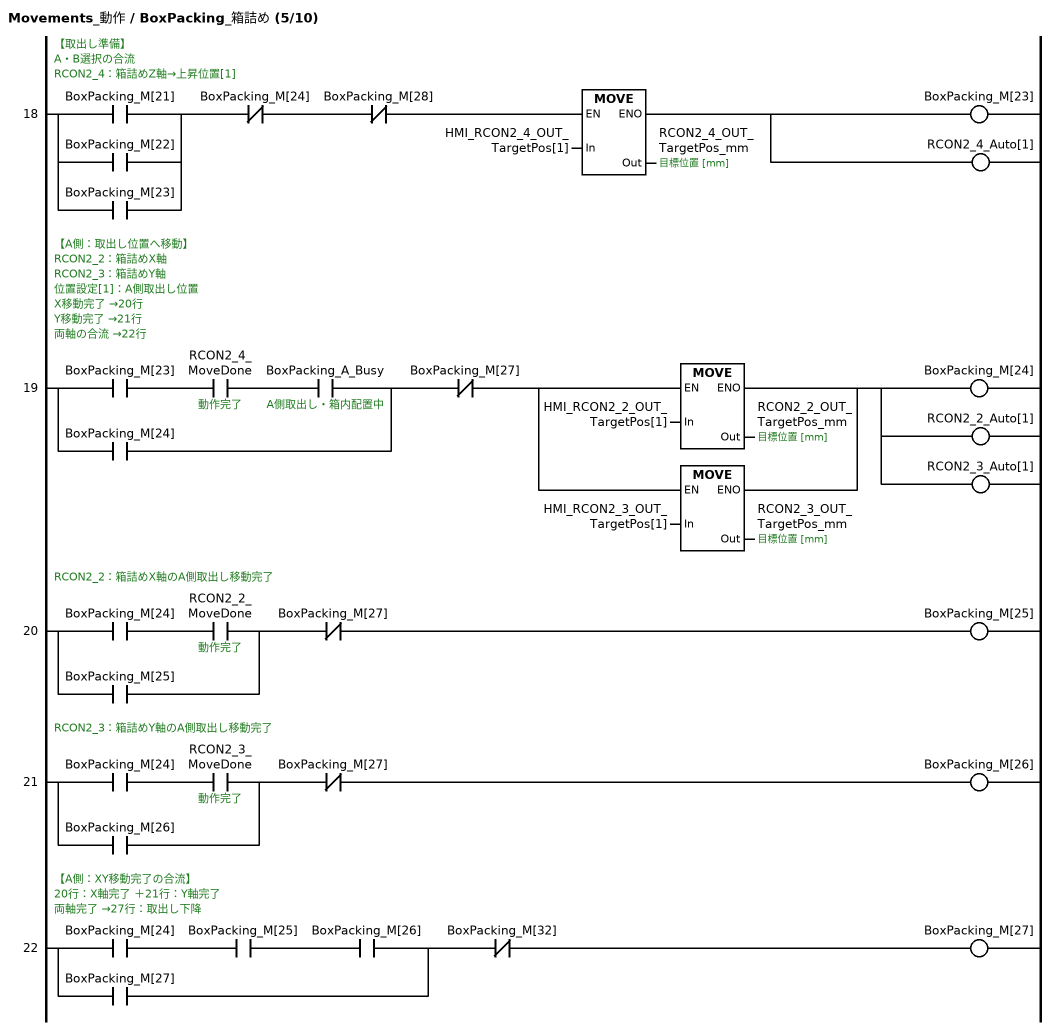
(* Rung 18: 【取出し準備】 / A・B選択の合流 / RCON2_4：箱詰めZ軸→上昇位置[1] *)
IF (BoxPacking_M[21] OR BoxPacking_M[22] OR BoxPacking_M[23]) AND NOT BoxPacking_M[24] AND NOT BoxPacking_M[28] THEN
    RCON2_4_OUT_TargetPos_mm := HMI_RCON2_4_OUT_TargetPos[1];
END_IF;
_p154 := (BoxPacking_M[21] OR BoxPacking_M[22] OR BoxPacking_M[23]) AND NOT BoxPacking_M[24] AND NOT BoxPacking_M[28];
BoxPacking_M[23] := _p154;
RCON2_4_Auto[1] := _p154;
(* Rung 19: 【A側：取出し位置へ移動】 / RCON2_2：箱詰めX軸 / RCON2_3：箱詰めY軸 / 位置設定[1]：A側取出し位置 / X移動完了 →20行 / Y移動完了 →21行 / 両軸の合流 →22行 *)
_p155 := ((BoxPacking_M[23] AND RCON2_4_MoveDone AND BoxPacking_A_Busy) OR BoxPacking_M[24]) AND NOT BoxPacking_M[27];
IF _p155 THEN
    RCON2_2_OUT_TargetPos_mm := HMI_RCON2_2_OUT_TargetPos[1];
    RCON2_3_OUT_TargetPos_mm := HMI_RCON2_3_OUT_TargetPos[1];
END_IF;
BoxPacking_M[24] := _p155;
RCON2_2_Auto[1] := _p155;
RCON2_3_Auto[1] := _p155;
(* Rung 20: RCON2_2：箱詰めX軸のA側取出し移動完了 *)
BoxPacking_M[25] := ((BoxPacking_M[24] AND RCON2_2_MoveDone) OR BoxPacking_M[25]) AND NOT BoxPacking_M[27];
(* Rung 21: RCON2_3：箱詰めY軸のA側取出し移動完了 *)
BoxPacking_M[26] := ((BoxPacking_M[24] AND RCON2_3_MoveDone) OR BoxPacking_M[26]) AND NOT BoxPacking_M[27];
(* Rung 22: 【A側：XY移動完了の合流】 / 20行：X軸完了 ＋21行：Y軸完了 / 両軸完了 →27行：取出し下降 *)
BoxPacking_M[27] := ((BoxPacking_M[24] AND BoxPacking_M[25] AND BoxPacking_M[26]) OR BoxPacking_M[27]) AND NOT BoxPacking_M[32];

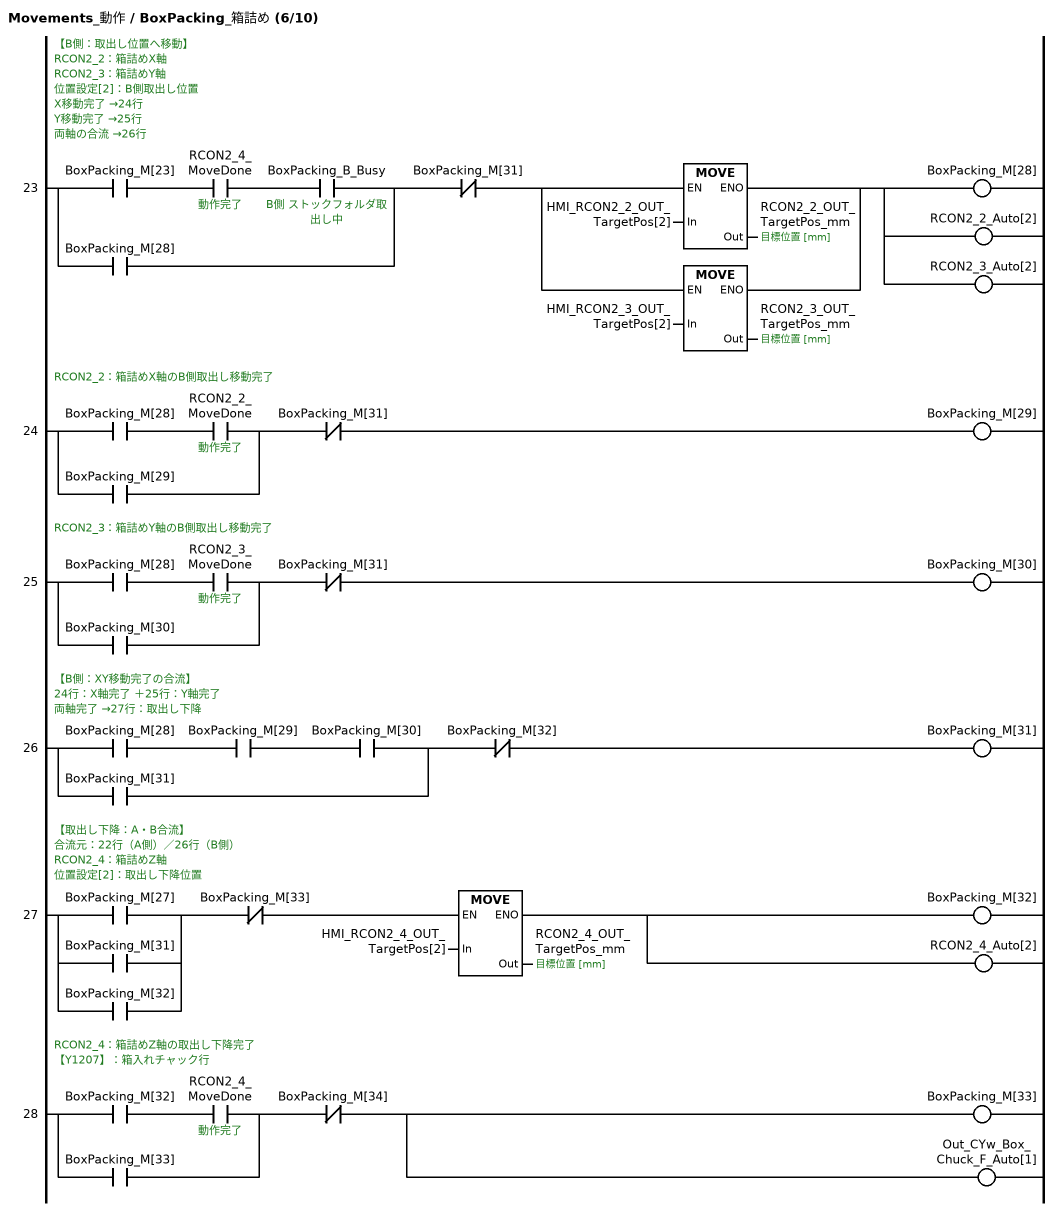
(* Rung 23: 【B側：取出し位置へ移動】 / RCON2_2：箱詰めX軸 / RCON2_3：箱詰めY軸 / 位置設定[2]：B側取出し位置 / X移動完了 →24行 / Y移動完了 →25行 / 両軸の合流 →26行 *)
_p156 := ((BoxPacking_M[23] AND RCON2_4_MoveDone AND BoxPacking_B_Busy) OR BoxPacking_M[28]) AND NOT BoxPacking_M[31];
IF _p156 THEN
    RCON2_2_OUT_TargetPos_mm := HMI_RCON2_2_OUT_TargetPos[2];
    RCON2_3_OUT_TargetPos_mm := HMI_RCON2_3_OUT_TargetPos[2];
END_IF;
BoxPacking_M[28] := _p156;
RCON2_2_Auto[2] := _p156;
RCON2_3_Auto[2] := _p156;
(* Rung 24: RCON2_2：箱詰めX軸のB側取出し移動完了 *)
BoxPacking_M[29] := ((BoxPacking_M[28] AND RCON2_2_MoveDone) OR BoxPacking_M[29]) AND NOT BoxPacking_M[31];
(* Rung 25: RCON2_3：箱詰めY軸のB側取出し移動完了 *)
BoxPacking_M[30] := ((BoxPacking_M[28] AND RCON2_3_MoveDone) OR BoxPacking_M[30]) AND NOT BoxPacking_M[31];
(* Rung 26: 【B側：XY移動完了の合流】 / 24行：X軸完了 ＋25行：Y軸完了 / 両軸完了 →27行：取出し下降 *)
BoxPacking_M[31] := ((BoxPacking_M[28] AND BoxPacking_M[29] AND BoxPacking_M[30]) OR BoxPacking_M[31]) AND NOT BoxPacking_M[32];
(* Rung 27: 【取出し下降：A・B合流】 / 合流元：22行（A側）／26行（B側） / RCON2_4：箱詰めZ軸 / 位置設定[2]：取出し下降位置 *)
IF (BoxPacking_M[27] OR BoxPacking_M[31] OR BoxPacking_M[32]) AND NOT BoxPacking_M[33] THEN
    RCON2_4_OUT_TargetPos_mm := HMI_RCON2_4_OUT_TargetPos[2];
END_IF;
_p157 := (BoxPacking_M[27] OR BoxPacking_M[31] OR BoxPacking_M[32]) AND NOT BoxPacking_M[33];
BoxPacking_M[32] := _p157;
RCON2_4_Auto[2] := _p157;
(* Rung 28: RCON2_4：箱詰めZ軸の取出し下降完了 / 【Y1207】：箱入れチャック行 *)
_p158 := ((BoxPacking_M[32] AND RCON2_4_MoveDone) OR BoxPacking_M[33]) AND NOT BoxPacking_M[34];
BoxPacking_M[33] := _p158;
Out_CYw_Box_Chuck_F_Auto[1] := _p158;

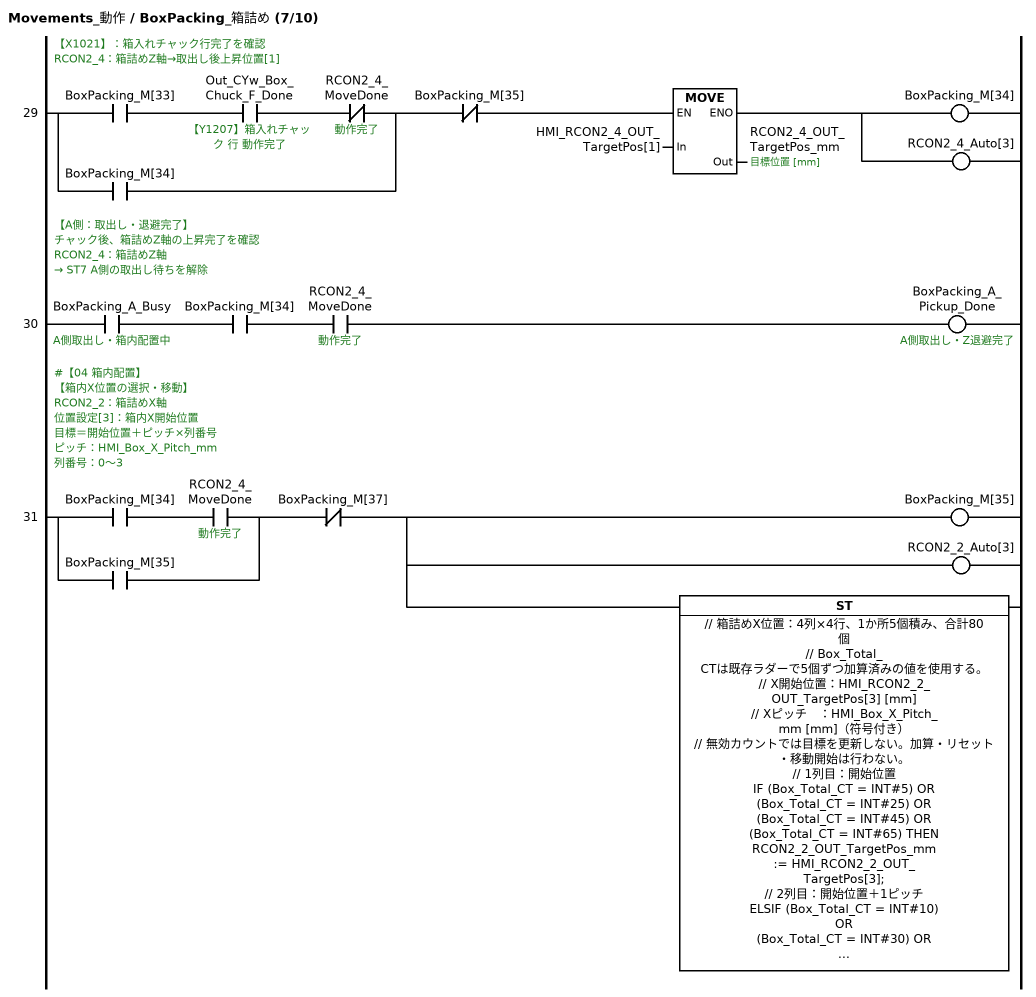
(* Rung 29: 【X1021】：箱入れチャック行完了を確認 / RCON2_4：箱詰めZ軸→取出し後上昇位置[1] *)
IF ((BoxPacking_M[33] AND Out_CYw_Box_Chuck_F_Done AND NOT RCON2_4_MoveDone) OR BoxPacking_M[34]) AND NOT BoxPacking_M[35] THEN
    RCON2_4_OUT_TargetPos_mm := HMI_RCON2_4_OUT_TargetPos[1];
END_IF;
_p159 := ((BoxPacking_M[33] AND Out_CYw_Box_Chuck_F_Done AND NOT RCON2_4_MoveDone) OR BoxPacking_M[34]) AND NOT BoxPacking_M[35];
BoxPacking_M[34] := _p159;
RCON2_4_Auto[3] := _p159;
(* Rung 30: 【A側：取出し・退避完了】 / チャック後、箱詰めZ軸の上昇完了を確認 / RCON2_4：箱詰めZ軸 / → ST7 A側の取出し待ちを解除 *)
BoxPacking_A_Pickup_Done := BoxPacking_A_Busy AND BoxPacking_M[34] AND RCON2_4_MoveDone;
(* Rung 31: #【04 箱内配置】 / 【箱内X位置の選択・移動】 / RCON2_2：箱詰めX軸 / 位置設定[3]：箱内X開始位置 / 目標＝開始位置＋ピッチ×列番号 / ピッチ：HMI_Box_X_Pitch_mm / 列番号：0～3 *)
_p160 := ((BoxPacking_M[34] AND RCON2_4_MoveDone) OR BoxPacking_M[35]) AND NOT BoxPacking_M[37];
BoxPacking_M[35] := _p160;
RCON2_2_Auto[3] := _p160;
IF _p160 THEN
    // 箱詰めX位置：4列×4行、1か所5個積み、合計80個
    // Box_Total_CTは既存ラダーで5個ずつ加算済みの値を使用する。
    // X開始位置：HMI_RCON2_2_OUT_TargetPos[3] [mm]
    // Xピッチ　：HMI_Box_X_Pitch_mm [mm]（符号付き）
    // 無効カウントでは目標を更新しない。加算・リセット・移動開始は行わない。
    
    // 1列目：開始位置
    IF (Box_Total_CT = INT#5) OR
       (Box_Total_CT = INT#25) OR
       (Box_Total_CT = INT#45) OR
       (Box_Total_CT = INT#65) THEN
    
        RCON2_2_OUT_TargetPos_mm := HMI_RCON2_2_OUT_TargetPos[3];
    
    // 2列目：開始位置＋1ピッチ
    ELSIF (Box_Total_CT = INT#10) OR
          (Box_Total_CT = INT#30) OR
          (Box_Total_CT = INT#50) OR
          (Box_Total_CT = INT#70) THEN
    
        RCON2_2_OUT_TargetPos_mm :=
            HMI_RCON2_2_OUT_TargetPos[3] +
            HMI_Box_X_Pitch_mm;
    
    // 3列目：開始位置＋2ピッチ
    ELSIF (Box_Total_CT = INT#15) OR
          (Box_Total_CT = INT#35) OR
          (Box_Total_CT = INT#55) OR
          (Box_Total_CT = INT#75) THEN
    
        RCON2_2_OUT_TargetPos_mm :=
            HMI_RCON2_2_OUT_TargetPos[3] +
            HMI_Box_X_Pitch_mm * LREAL#2.0;
    
    // 4列目：開始位置＋3ピッチ
    ELSIF (Box_Total_CT = INT#20) OR
          (Box_Total_CT = INT#40) OR
          (Box_Total_CT = INT#60) OR
          (Box_Total_CT = INT#80) THEN
    
        RCON2_2_OUT_TargetPos_mm :=
            HMI_RCON2_2_OUT_TargetPos[3] +
            HMI_Box_X_Pitch_mm * LREAL#3.0;
    END_IF;
END_IF;

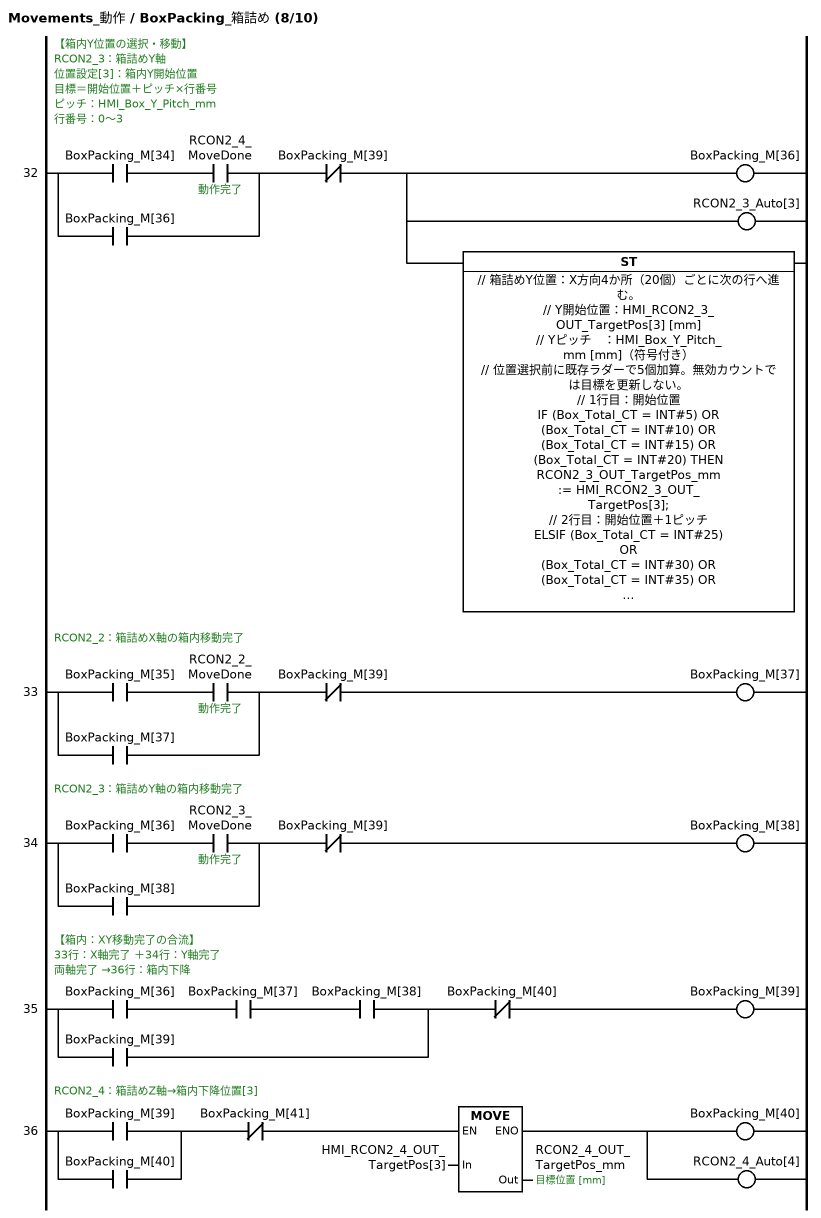
(* Rung 32: 【箱内Y位置の選択・移動】 / RCON2_3：箱詰めY軸 / 位置設定[3]：箱内Y開始位置 / 目標＝開始位置＋ピッチ×行番号 / ピッチ：HMI_Box_Y_Pitch_mm / 行番号：0～3 *)
_p161 := ((BoxPacking_M[34] AND RCON2_4_MoveDone) OR BoxPacking_M[36]) AND NOT BoxPacking_M[39];
BoxPacking_M[36] := _p161;
RCON2_3_Auto[3] := _p161;
IF _p161 THEN
    // 箱詰めY位置：X方向4か所（20個）ごとに次の行へ進む。
    // Y開始位置：HMI_RCON2_3_OUT_TargetPos[3] [mm]
    // Yピッチ　：HMI_Box_Y_Pitch_mm [mm]（符号付き）
    // 位置選択前に既存ラダーで5個加算。無効カウントでは目標を更新しない。
    
    // 1行目：開始位置
    IF (Box_Total_CT = INT#5) OR
       (Box_Total_CT = INT#10) OR
       (Box_Total_CT = INT#15) OR
       (Box_Total_CT = INT#20) THEN
    
        RCON2_3_OUT_TargetPos_mm := HMI_RCON2_3_OUT_TargetPos[3];
    
    // 2行目：開始位置＋1ピッチ
    ELSIF (Box_Total_CT = INT#25) OR
          (Box_Total_CT = INT#30) OR
          (Box_Total_CT = INT#35) OR
          (Box_Total_CT = INT#40) THEN
    
        RCON2_3_OUT_TargetPos_mm :=
            HMI_RCON2_3_OUT_TargetPos[3] + HMI_Box_Y_Pitch_mm;
    
    // 3行目：開始位置＋2ピッチ
    ELSIF (Box_Total_CT = INT#45) OR
          (Box_Total_CT = INT#50) OR
          (Box_Total_CT = INT#55) OR
          (Box_Total_CT = INT#60) THEN
    
        RCON2_3_OUT_TargetPos_mm :=
            HMI_RCON2_3_OUT_TargetPos[3] + HMI_Box_Y_Pitch_mm * LREAL#2.0;
    
    // 4行目：開始位置＋3ピッチ
    ELSIF (Box_Total_CT = INT#65) OR
          (Box_Total_CT = INT#70) OR
          (Box_Total_CT = INT#75) OR
          (Box_Total_CT = INT#80) THEN
    
        RCON2_3_OUT_TargetPos_mm :=
            HMI_RCON2_3_OUT_TargetPos[3] + HMI_Box_Y_Pitch_mm * LREAL#3.0;
    END_IF;
END_IF;
(* Rung 33: RCON2_2：箱詰めX軸の箱内移動完了 *)
BoxPacking_M[37] := ((BoxPacking_M[35] AND RCON2_2_MoveDone) OR BoxPacking_M[37]) AND NOT BoxPacking_M[39];
(* Rung 34: RCON2_3：箱詰めY軸の箱内移動完了 *)
BoxPacking_M[38] := ((BoxPacking_M[36] AND RCON2_3_MoveDone) OR BoxPacking_M[38]) AND NOT BoxPacking_M[39];
(* Rung 35: 【箱内：XY移動完了の合流】 / 33行：X軸完了 ＋34行：Y軸完了 / 両軸完了 →36行：箱内下降 *)
BoxPacking_M[39] := ((BoxPacking_M[36] AND BoxPacking_M[37] AND BoxPacking_M[38]) OR BoxPacking_M[39]) AND NOT BoxPacking_M[40];
(* Rung 36: RCON2_4：箱詰めZ軸→箱内下降位置[3] *)
IF (BoxPacking_M[39] OR BoxPacking_M[40]) AND NOT BoxPacking_M[41] THEN
    RCON2_4_OUT_TargetPos_mm := HMI_RCON2_4_OUT_TargetPos[3];
END_IF;
_p162 := (BoxPacking_M[39] OR BoxPacking_M[40]) AND NOT BoxPacking_M[41];
BoxPacking_M[40] := _p162;
RCON2_4_Auto[4] := _p162;

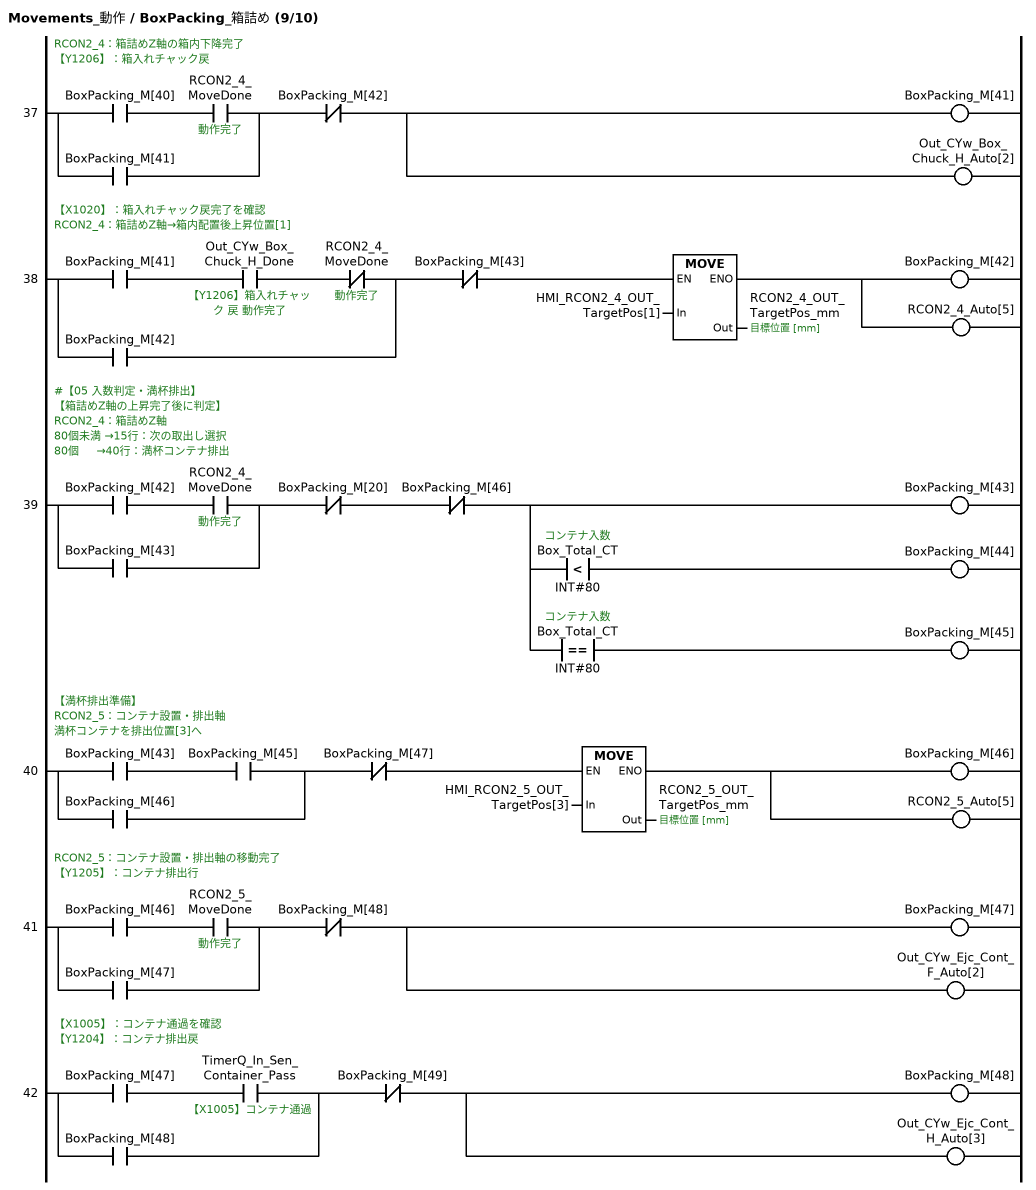
(* Rung 37: RCON2_4：箱詰めZ軸の箱内下降完了 / 【Y1206】：箱入れチャック戻 *)
_p163 := ((BoxPacking_M[40] AND RCON2_4_MoveDone) OR BoxPacking_M[41]) AND NOT BoxPacking_M[42];
BoxPacking_M[41] := _p163;
Out_CYw_Box_Chuck_H_Auto[2] := _p163;
(* Rung 38: 【X1020】：箱入れチャック戻完了を確認 / RCON2_4：箱詰めZ軸→箱内配置後上昇位置[1] *)
IF ((BoxPacking_M[41] AND Out_CYw_Box_Chuck_H_Done AND NOT RCON2_4_MoveDone) OR BoxPacking_M[42]) AND NOT BoxPacking_M[43] THEN
    RCON2_4_OUT_TargetPos_mm := HMI_RCON2_4_OUT_TargetPos[1];
END_IF;
_p164 := ((BoxPacking_M[41] AND Out_CYw_Box_Chuck_H_Done AND NOT RCON2_4_MoveDone) OR BoxPacking_M[42]) AND NOT BoxPacking_M[43];
BoxPacking_M[42] := _p164;
RCON2_4_Auto[5] := _p164;
(* Rung 39: #【05 入数判定・満杯排出】 / 【箱詰めZ軸の上昇完了後に判定】 / RCON2_4：箱詰めZ軸 / 80個未満 →15行：次の取出し選択 / 80個     →40行：満杯コンテナ排出 *)
_p165 := ((BoxPacking_M[42] AND RCON2_4_MoveDone) OR BoxPacking_M[43]) AND NOT BoxPacking_M[20] AND NOT BoxPacking_M[46];
BoxPacking_M[43] := _p165;
BoxPacking_M[44] := _p165 AND (Box_Total_CT < INT#80);
BoxPacking_M[45] := _p165 AND (Box_Total_CT = INT#80);
(* Rung 40: 【満杯排出準備】 / RCON2_5：コンテナ設置・排出軸 / 満杯コンテナを排出位置[3]へ *)
IF ((BoxPacking_M[43] AND BoxPacking_M[45]) OR BoxPacking_M[46]) AND NOT BoxPacking_M[47] THEN
    RCON2_5_OUT_TargetPos_mm := HMI_RCON2_5_OUT_TargetPos[3];
END_IF;
_p166 := ((BoxPacking_M[43] AND BoxPacking_M[45]) OR BoxPacking_M[46]) AND NOT BoxPacking_M[47];
BoxPacking_M[46] := _p166;
RCON2_5_Auto[5] := _p166;
(* Rung 41: RCON2_5：コンテナ設置・排出軸の移動完了 / 【Y1205】：コンテナ排出行 *)
_p167 := ((BoxPacking_M[46] AND RCON2_5_MoveDone) OR BoxPacking_M[47]) AND NOT BoxPacking_M[48];
BoxPacking_M[47] := _p167;
Out_CYw_Ejc_Cont_F_Auto[2] := _p167;
(* Rung 42: 【X1005】：コンテナ通過を確認 / 【Y1204】：コンテナ排出戻 *)
_p168 := ((BoxPacking_M[47] AND TimerQ_In_Sen_Container_Pass) OR BoxPacking_M[48]) AND NOT BoxPacking_M[49];
BoxPacking_M[48] := _p168;
Out_CYw_Ejc_Cont_H_Auto[3] := _p168;

